METHOD PRIVATE parseFaults : BOOL
VAR
    _q  : UDINT;
    _s  : UDINT;
END_VAR
_q := _device.DCMeter.DCQuesReg;
_s := _swFaultReg;

IF ITECH_Type = 'IT6600C' THEN
    _DeviceFaults.overVoltageProtection  := _q.0;
    _DeviceFaults.overCurrentProtection  := _q.1;
    _DeviceFaults.overPowerProtection    := _q.2;
    _DeviceFaults.underVoltageProtection := _q.3;
    _DeviceFaults.overTempProtection     := _q.4;
    _DeviceFaults.underCurrentProtection := _q.5;
    _DeviceFaults.senseFault             := _q.6;
    _DeviceFaults.currentSharingFault    := _q.7;
    _DeviceFaults.externalInhibit        := _q.9;
    _DeviceFaults.faultProtection        := _q.10;
    _DeviceFaults.loopOscFailure         := _q.11;
    _DeviceFaults.outputNotRegulated     := _q.12;

    _SoftwareFaults.overVoltageProtection         := _s.0;
    _SoftwareFaults.positiveOverCurrentProtection := _s.1;
    _SoftwareFaults.negativeOverCurrentProtection := _s.2;
    _SoftwareFaults.positiveOverPowerProtection   := _s.3;
    _SoftwareFaults.negativeOverPowerProtection   := _s.4;
    _SoftwareFaults.underCurrentProtection        := _s.5;
    _SoftwareFaults.underVoltageProtection        := _s.6;
    _SoftwareFaults.overTemperatureProtection     := _s.7;
END_IF

IF ITECH_Type = 'IT6000' THEN
    _DeviceFaults.overVoltageProtection  := _q.0;
    _DeviceFaults.overCurrentProtection  := _q.1 OR _q.2;
    _DeviceFaults.overPowerProtection    := _q.3 OR _q.4;
    _DeviceFaults.underVoltageProtection := _q.5;
    _DeviceFaults.overTempProtection     := _q.6;
    _DeviceFaults.underCurrentProtection := _q.7;
    _DeviceFaults.senseFault             := _q.8;
    _DeviceFaults.currentSharingFault    := _q.9;
    // bit 10: output reversed (reported through the software-fault register instead)
    _DeviceFaults.externalInhibit        := _q.11;
    _DeviceFaults.faultProtection        := _q.12;
    _DeviceFaults.loopOscFailure         := _q.13;
END_IF

_SoftwareFaults.senseAbnormal                     := _s.8;
_SoftwareFaults.senseReverseProtection            := _s.9;
_SoftwareFaults.outputReverseProtection           := _s.10;
_SoftwareFaults.multiMasterUnitsAbnormal          := _s.11;
_SoftwareFaults.opticalFiberUnlocked_multiMaster  := _s.12;
_SoftwareFaults.opticalFiberUnlocked_singleMaster := _s.13;
_SoftwareFaults.moduleCheckingFailure             := _s.14;
_SoftwareFaults.unevenCurrentProtection           := _s.15;
_SoftwareFaults.hardwareProtection                := _s.16;
_SoftwareFaults.masterUnitPowerFailureProtection  := _s.17;
_SoftwareFaults.inhibit_latchmode                 := _s.18;
_SoftwareFaults.inhibit_livingMode                := _s.19;
_SoftwareFaults.capacitorOverCurrentprotection    := _s.20;
_SoftwareFaults.slaveUnitPowerFailureProtection   := _s.21;
END_METHOD

METHOD PRIVATE rdReal : REAL
VAR_INPUT
    inpIdx      : UINT;
    inpKeep     : REAL;     // returned unchanged unless this signal's last read was good
END_VAR
IF inpIdx <= _readCount AND _arrReadResults[inpIdx].quality = E_SignalQuality.Good THEN
    rdReal := _arrReadResults[inpIdx].valueReal;
ELSE
    rdReal := inpKeep;
END_IF
END_METHOD

METHOD PRIVATE rdUdint : UDINT
VAR_INPUT
    inpIdx      : UINT;
    inpKeep     : UDINT;
END_VAR
IF inpIdx <= _readCount AND _arrReadResults[inpIdx].quality = E_SignalQuality.Good THEN
    rdUdint := _arrReadResults[inpIdx].valueUdint;
ELSE
    rdUdint := inpKeep;
END_IF
END_METHOD

METHOD PRIVATE readImage : BOOL
_device.DCMeter.DCVrms     := rdReal(cRD_METER + 1, _device.DCMeter.DCVrms);
_device.DCMeter.DCIrms     := rdReal(cRD_METER + 2, _device.DCMeter.DCIrms);
_device.DCMeter.DCPrms     := rdReal(cRD_METER + 3, _device.DCMeter.DCPrms);
_device.DCMeter.DCOperReg  := rdUdint(cRD_METER + 4, _device.DCMeter.DCOperReg);
_device.DCMeter.DCStateReg := rdUdint(cRD_METER + 5, _device.DCMeter.DCStateReg);
_device.DCMeter.DCQuesReg  := rdUdint(cRD_METER + 6, _device.DCMeter.DCQuesReg);

_device.DCSource.DCMode          := rdUdint(cRD_SOURCE + 1,  _device.DCSource.DCMode);
_device.DCSource.DCVoltSP        := rdReal(cRD_SOURCE + 2,   _device.DCSource.DCVoltSP);
_device.DCSource.DCVoltRise      := rdReal(cRD_SOURCE + 3,   _device.DCSource.DCVoltRise);
_device.DCSource.DCVoltFall      := rdReal(cRD_SOURCE + 4,   _device.DCSource.DCVoltFall);
_device.DCSource.DCCurrentSP     := rdReal(cRD_SOURCE + 5,   _device.DCSource.DCCurrentSP);
_device.DCSource.DCCurrentRise   := rdReal(cRD_SOURCE + 6,   _device.DCSource.DCCurrentRise);
_device.DCSource.DCCurrentFall   := rdReal(cRD_SOURCE + 7,   _device.DCSource.DCCurrentFall);
_device.DCSource.DCVoltHigh      := rdReal(cRD_SOURCE + 8,   _device.DCSource.DCVoltHigh);
_device.DCSource.DCVoltLow       := rdReal(cRD_SOURCE + 9,   _device.DCSource.DCVoltLow);
_device.DCSource.DCCurrentHigh   := rdReal(cRD_SOURCE + 10,  _device.DCSource.DCCurrentHigh);
_device.DCSource.DCCurrentLow    := rdReal(cRD_SOURCE + 11,  _device.DCSource.DCCurrentLow);
_device.DCSource.DCCC_SpeedState := rdUdint(cRD_SOURCE + 12, _device.DCSource.DCCC_SpeedState);
_device.DCSource.DCCV_SpeedState := rdUdint(cRD_SOURCE + 13, _device.DCSource.DCCV_SpeedState);
_device.DCSource.DCPowerHigh     := rdReal(cRD_SOURCE + 14,  _device.DCSource.DCPowerHigh);
_device.DCSource.DCPowerLow      := rdReal(cRD_SOURCE + 15,  _device.DCSource.DCPowerLow);

_device.Protection.OVPState  := rdUdint(cRD_PROT + 1,  _device.Protection.OVPState);
_device.Protection.OVPLevel  := rdReal(cRD_PROT + 2,   _device.Protection.OVPLevel);
_device.Protection.OVPDelay  := rdReal(cRD_PROT + 3,   _device.Protection.OVPDelay);
_device.Protection.OCPState  := rdUdint(cRD_PROT + 4,  _device.Protection.OCPState);
_device.Protection.OCPLevel  := rdReal(cRD_PROT + 5,   _device.Protection.OCPLevel);
_device.Protection.OCPDelay  := rdReal(cRD_PROT + 6,   _device.Protection.OCPDelay);
_device.Protection.OPPState  := rdUdint(cRD_PROT + 7,  _device.Protection.OPPState);
_device.Protection.OPPLevel  := rdReal(cRD_PROT + 8,   _device.Protection.OPPLevel);
_device.Protection.OPPDelay  := rdReal(cRD_PROT + 9,   _device.Protection.OPPDelay);
_device.Protection.UCPState  := rdUdint(cRD_PROT + 10, _device.Protection.UCPState);
_device.Protection.UCPLevel  := rdReal(cRD_PROT + 11,  _device.Protection.UCPLevel);
_device.Protection.UCPDelay  := rdReal(cRD_PROT + 12,  _device.Protection.UCPDelay);
_device.Protection.UCPWarmup := rdReal(cRD_PROT + 13,  _device.Protection.UCPWarmup);
_device.Protection.UVPState  := rdUdint(cRD_PROT + 14, _device.Protection.UVPState);
_device.Protection.UVPLevel  := rdReal(cRD_PROT + 15,  _device.Protection.UVPLevel);
_device.Protection.UVPDelay  := rdReal(cRD_PROT + 16,  _device.Protection.UVPDelay);
_device.Protection.UVPWarmup := rdReal(cRD_PROT + 17,  _device.Protection.UVPWarmup);

_swFaultReg := rdUdint(cRD_SWF, _swFaultReg);

_device.System.ON_OFF            := rdUdint(cRD_SYS + 1, _device.System.ON_OFF);
_device.System.SenseVolt         := rdReal(cRD_SYS + 2,  _device.System.SenseVolt);
_device.System.Heartbeat         := rdUdint(cRD_SYS + 3, _device.System.Heartbeat);
_device.System.Timer_ON_OFF      := rdUdint(cRD_SYS + 4, _device.System.Timer_ON_OFF);
_device.System.RemoteSenseStatus := rdUdint(cRD_SYS + 5, _device.System.RemoteSenseStatus);
_device.System.RemoteSenseLevel  := rdReal(cRD_SYS + 6,  _device.System.RemoteSenseLevel);
_device.System.OutputRZero       := rdUdint(cRD_SYS + 7, _device.System.OutputRZero);
_device.System.MeasureCycle      := rdUdint(cRD_SYS + 8, _device.System.MeasureCycle);
END_METHOD

METHOD PRIVATE runComms : BOOL
VAR
    _i      : UINT;
END_VAR
// A reset (rising edge) re-arms comms and queues the supply's own protection reset.
_resetTrig(CLK := _resetCalled);
_resetCalled := FALSE;
IF _resetTrig.Q THEN
    _commFaulted := FALSE;
    _deviceResetPending := TRUE;
END_IF

// A type change while running takes comms down for one scan so the driver re-reads its tables.
_mapChanged := _commRunPrev AND (ITECH_Type <> _activeType);
_commRun := _enabled AND _mapValid AND NOT _commFaulted AND NOT _mapChanged;

IF _commRun AND NOT _commRunPrev THEN
    configureDriver();
    _baselineTaken  := FALSE;
    _lastReadCycles := 0;
    _tonReadWatchdog(IN := FALSE);
END_IF
_commRunPrev := _commRun;

IF _baselineTaken THEN
    writeImage();
END_IF

_mb(
    inpEnable           := _commRun,
    inpHoldWrites       := NOT _baselineTaken,
    inpPtrReadConfig    := ADR(_arrReadConfig),
    inpPtrWriteConfig   := ADR(_arrWriteConfig),
    inpPtrReadResults   := ADR(_arrReadResults),
    inpPtrWriteData     := ADR(_arrWriteData));
_mb.cycle();

IF NOT _commRun THEN
    _tonReadWatchdog(IN := FALSE);
    deviceResetWrite();         // keeps the one-shot driver disabled
    RETURN;
END_IF

// ── the latch: the FIRST failed transaction stops everything ────────────────────────────────
IF _mb.stsError THEN
    latchCommFault('Modbus driver configuration error - comms stopped until reset');
    RETURN;
END_IF
FOR _i := 1 TO _readCount DO
    IF _arrReadResults[_i].quality = E_SignalQuality.BadComm THEN
        latchCommFault('Modbus read failed - comms stopped until reset');
        RETURN;
    END_IF
END_FOR
FOR _i := 1 TO cWR_PROT + 17 DO
    IF _arrWriteData[_i].writeError THEN
        latchCommFault('Modbus write failed - comms stopped until reset');
        RETURN;
    END_IF
END_FOR

// A driver that stops completing read cycles without reporting an error is a fault too.
IF _mb.stsStatus.totalReadCycles <> _lastReadCycles THEN
    _lastReadCycles := _mb.stsStatus.totalReadCycles;
    _tonReadWatchdog(IN := FALSE);
END_IF
_tonReadWatchdog(IN := TRUE, PT := _wdTime);
IF _tonReadWatchdog.Q THEN
    latchCommFault('Modbus read watchdog: no read cycle completed - comms stopped until reset');
    RETURN;
END_IF

readImage();

// First complete, clean read cycle since (re)start: seed the command image from the supply,
// then release writes.
IF NOT _baselineTaken AND _mb.stsStatus.totalReadCycles > 0 THEN
    _command := _device;
    IF _baselineCurrentLimit > 0 THEN
        cmdSetCurrentLimits(currentLimitHigh := _baselineCurrentLimit,
                            currentLimitLow  := -_baselineCurrentLimit);
    END_IF
    initParameters();
    IF _commFaultSeen THEN
        cmdDCSourceEnable(FALSE);       // also zeroes the operator's ON/OFF request
        _commFaultSeen := FALSE;
    END_IF
    _baselineTaken := TRUE;
END_IF

deviceResetWrite();
END_METHOD

METHOD PRIVATE selectRegisterMap : BOOL
_mapValid := TRUE;

IF ITECH_Type = 'IT6600C' THEN
    _regDCMeter         := 1401;
    _regDCSource        := 1201;
    _regSystemStatus    := 1001;
    _regProtection      := 1701;
    _regSoftwareFaults  := 1803;
    _regOnOff           := 1001;
    _regResetFault      := 1801;
    _scanTime           := T#100MS;
    _hasExtStatus       := TRUE;
ELSIF ITECH_Type = 'IT6000' THEN
    _regDCMeter         := 1107;
    _regDCSource        := 1019;
    _regSystemStatus    := 1001;
    _regProtection      := 1169;
    _regSoftwareFaults  := 1225;
    _regOnOff           := 1001;
    _regResetFault      := 1223;
    _scanTime           := T#250MS;
    _hasExtStatus       := FALSE;
ELSE
    _mapValid := FALSE;
END_IF
END_METHOD

METHOD setCommandValues : BOOL
IF NOT inpAuto THEN
    IF NOT stsFaulted THEN
        _command.System.ON_OFF     := HMI_DeviceSignals.deviceSignals_write.System.ON_OFF;
        _command.DCSource.DCMode   := HMI_DeviceSignals.deviceSignals_write.DCSource.DCMode;
    END_IF
    _command.DCSource.DCPowerHigh   := HMI_DeviceSignals.deviceSignals_write.DCSource.DCPowerHigh;
    _command.DCSource.DCPowerLow    := HMI_DeviceSignals.deviceSignals_write.DCSource.DCPowerLow;
    _command.DCSource.DCCurrentSP   := HMI_DeviceSignals.deviceSignals_write.DCSource.DCCurrentSP;
    _command.DCSource.DCCurrentRise := HMI_DeviceSignals.deviceSignals_write.DCSource.DCCurrentRise;
    _command.DCSource.DCCurrentFall := HMI_DeviceSignals.deviceSignals_write.DCSource.DCCurrentFall;
    _command.DCSource.DCCurrentHigh := HMI_DeviceSignals.deviceSignals_write.DCSource.DCCurrentHigh;
    _command.DCSource.DCCurrentLow  := HMI_DeviceSignals.deviceSignals_write.DCSource.DCCurrentLow;
    _command.DCSource.DCVoltSP      := HMI_DeviceSignals.deviceSignals_write.DCSource.DCVoltSP;
    _command.DCSource.DCVoltRise    := HMI_DeviceSignals.deviceSignals_write.DCSource.DCVoltRise;
    _command.DCSource.DCVoltFall    := HMI_DeviceSignals.deviceSignals_write.DCSource.DCVoltFall;
    _command.DCSource.DCVoltHigh    := HMI_DeviceSignals.deviceSignals_write.DCSource.DCVoltHigh;
    _command.DCSource.DCVoltLow     := HMI_DeviceSignals.deviceSignals_write.DCSource.DCVoltLow;

    _command.Protection.OCPState    := HMI_DeviceSignals.deviceSignals_write.Protection.OCPState;
    _command.Protection.OCPLevel    := HMI_DeviceSignals.deviceSignals_write.Protection.OCPLevel;
    _command.Protection.OCPDelay    := HMI_DeviceSignals.deviceSignals_write.Protection.OCPDelay;
    _command.Protection.OVPState    := HMI_DeviceSignals.deviceSignals_write.Protection.OVPState;
    _command.Protection.OVPLevel    := HMI_DeviceSignals.deviceSignals_write.Protection.OVPLevel;
    _command.Protection.OVPDelay    := HMI_DeviceSignals.deviceSignals_write.Protection.OVPDelay;
    _command.Protection.UCPState    := HMI_DeviceSignals.deviceSignals_write.Protection.UCPState;
    _command.Protection.UCPLevel    := HMI_DeviceSignals.deviceSignals_write.Protection.UCPLevel;
    _command.Protection.UCPDelay    := HMI_DeviceSignals.deviceSignals_write.Protection.UCPDelay;
    _command.Protection.UVPState    := HMI_DeviceSignals.deviceSignals_write.Protection.UVPState;
    _command.Protection.UVPLevel    := HMI_DeviceSignals.deviceSignals_write.Protection.UVPLevel;
    _command.Protection.UVPDelay    := HMI_DeviceSignals.deviceSignals_write.Protection.UVPDelay;
    _command.Protection.OPPState    := HMI_DeviceSignals.deviceSignals_write.Protection.OPPState;
    _command.Protection.OPPLevel    := HMI_DeviceSignals.deviceSignals_write.Protection.OPPLevel;
    _command.Protection.OPPDelay    := HMI_DeviceSignals.deviceSignals_write.Protection.OPPDelay;
END_IF
END_METHOD

METHOD setConfigs : BOOL
VAR_INPUT
    configs : ST_ITECH_SetConfigs;
END_VAR
_command.DCSource.DCMode         := configs.dcSource.DCMode;
_command.DCSource.DCPowerHigh    := configs.dcSource.DCPowerHigh;
_command.DCSource.DCPowerLow     := configs.dcSource.DCPowerLow;
_command.DCSource.DCCurrentSP    := configs.dcSource.DCCurrentSP;
_command.DCSource.DCCurrentRise  := configs.dcSource.DCCurrentRise;
_command.DCSource.DCCurrentFall  := configs.dcSource.DCCurrentFall;
_command.DCSource.DCCurrentHigh  := configs.dcSource.DCCurrentHigh;
_command.DCSource.DCCurrentLow   := configs.dcSource.DCCurrentLow;
_command.DCSource.DCVoltSP       := configs.dcSource.DCVoltSP;
_command.DCSource.DCVoltRise     := configs.dcSource.DCVoltRise;
_command.DCSource.DCVoltFall     := configs.dcSource.DCVoltFall;
_command.DCSource.DCVoltHigh     := configs.dcSource.DCVoltHigh;
_command.DCSource.DCVoltLow      := configs.dcSource.DCVoltLow;

_command.Protection.OCPLevel     := configs.protection.OCPLevel;
_command.Protection.OCPDelay     := configs.protection.OCPDelay;
_command.Protection.UCPLevel     := configs.protection.UCPLevel;
_command.Protection.UCPDelay     := configs.protection.UCPDelay;
_command.Protection.OVPLevel     := configs.protection.OVPLevel;
_command.Protection.OVPDelay     := configs.protection.OVPDelay;
_command.Protection.UVPLevel     := configs.protection.UVPLevel;
_command.Protection.UVPDelay     := configs.protection.UVPDelay;
_command.Protection.OPPLevel     := configs.protection.OPPLevel;
_command.Protection.OPPDelay     := configs.protection.OPPDelay;

_command.Protection.UCPState     := configs.protection.UCPState;
_command.Protection.UVPState     := configs.protection.UVPState;
_command.Protection.OCPState     := configs.protection.OCPState;
_command.Protection.OVPState     := configs.protection.OVPState;
_command.Protection.OPPState     := configs.protection.OPPState;
END_METHOD

METHOD setInterlock : BOOL
Interlock.name := _DeviceName;
Interlock(inpConfig := _dataInterlock);
END_METHOD

METHOD PRIVATE setRead : BOOL
VAR_INPUT
    inpIdx      : UINT;
    inpReg      : UINT;     // protocol (0-based) holding-register address
    inpIsReal   : BOOL;     // TRUE = 32-bit float, FALSE = 32-bit unsigned
END_VAR
_arrReadConfig[inpIdx].modbusAddr := 400001 + UINT_TO_UDINT(inpReg);
IF inpIsReal THEN
    _arrReadConfig[inpIdx].dataType := E_MBDataType.mbReal32;
ELSE
    _arrReadConfig[inpIdx].dataType := E_MBDataType.mbUInt32;
END_IF
END_METHOD

METHOD setStatusValues : BOOL
stsDCSourceState := _device.System.ON_OFF;
stsDCMode        := _device.DCSource.DCMode;
stsDCSource_V_SP := _device.DCSource.DCVoltSP;
stsDCMeterV      := _device.DCMeter.DCVrms;
stsDCMeterI      := _device.DCMeter.DCIrms;
stsDCMeterP      := _device.DCMeter.DCPrms;
sendLog(CONCAT('DC Source state changed to ', TO_STRING(stsDCSourceState)), 1);
sendLog(CONCAT('DC Source Voltage setpoint set to ', TO_STRING(stsDCSource_V_SP)), 2);
sendLog(CONCAT('DC Source mode set to ', TO_STRING(stsDCMode)), 3);
END_METHOD

METHOD PRIVATE setWrite : BOOL
VAR_INPUT
    inpIdx      : UINT;
    inpReg      : UINT;
    inpIsReal   : BOOL;
END_VAR
_arrWriteConfig[inpIdx].modbusAddr := 400001 + UINT_TO_UDINT(inpReg);
IF inpIsReal THEN
    _arrWriteConfig[inpIdx].dataType := E_MBDataType.mbReal32;
ELSE
    _arrWriteConfig[inpIdx].dataType := E_MBDataType.mbUInt32;
END_IF
END_METHOD

METHOD PRIVATE updateHMI : BOOL
HMI_DeviceSignals.deviceSignals_read := _device;
END_METHOD

METHOD PRIVATE writeImage : BOOL
// ON/OFF goes out as two 16-bit registers, LOW word first — exactly the bytes the previous
// implementation sent (it wrote the raw UDINT, not the word-swapped image every other value
// uses). Kept byte-for-byte because the supplies run on it; it is the one asymmetry with the
// read side (which takes the register pair high word first), so verify against the supply's
// manual before "fixing" it.
_arrWriteData[cWR_ONOFF + 1].valueUint := UDINT_TO_UINT(_command.System.ON_OFF AND 16#FFFF);
_arrWriteData[cWR_ONOFF + 2].valueUint := UDINT_TO_UINT(SHR(_command.System.ON_OFF, 16));

// IT6000 power values are in kW, IT6600C power values in W
_arrWriteData[cWR_SOURCE + 1].valueUdint := _command.DCSource.DCMode;
_arrWriteData[cWR_SOURCE + 2].valueReal  := _command.DCSource.DCVoltSP;
_arrWriteData[cWR_SOURCE + 3].valueReal  := _command.DCSource.DCVoltRise;
_arrWriteData[cWR_SOURCE + 4].valueReal  := _command.DCSource.DCVoltFall;
_arrWriteData[cWR_SOURCE + 5].valueReal  := _command.DCSource.DCCurrentSP;
_arrWriteData[cWR_SOURCE + 6].valueReal  := _command.DCSource.DCCurrentRise;
_arrWriteData[cWR_SOURCE + 7].valueReal  := _command.DCSource.DCCurrentFall;
_arrWriteData[cWR_SOURCE + 8].valueReal  := _command.DCSource.DCVoltHigh;
_arrWriteData[cWR_SOURCE + 9].valueReal  := _command.DCSource.DCVoltLow;
_arrWriteData[cWR_SOURCE + 10].valueReal := _command.DCSource.DCCurrentHigh;
_arrWriteData[cWR_SOURCE + 11].valueReal := _command.DCSource.DCCurrentLow;
_arrWriteData[cWR_SOURCE + 12].valueUdint := _command.DCSource.DCCC_SpeedState;
_arrWriteData[cWR_SOURCE + 13].valueUdint := _command.DCSource.DCCV_SpeedState;
_arrWriteData[cWR_SOURCE + 14].valueReal := _command.DCSource.DCPowerHigh;
_arrWriteData[cWR_SOURCE + 15].valueReal := _command.DCSource.DCPowerLow;

_arrWriteData[cWR_PROT + 1].valueUdint  := _command.Protection.OVPState;
_arrWriteData[cWR_PROT + 2].valueReal   := _command.Protection.OVPLevel;
_arrWriteData[cWR_PROT + 3].valueReal   := _command.Protection.OVPDelay;
_arrWriteData[cWR_PROT + 4].valueUdint  := _command.Protection.OCPState;
_arrWriteData[cWR_PROT + 5].valueReal   := _command.Protection.OCPLevel;
_arrWriteData[cWR_PROT + 6].valueReal   := _command.Protection.OCPDelay;
_arrWriteData[cWR_PROT + 7].valueUdint  := _command.Protection.OPPState;
_arrWriteData[cWR_PROT + 8].valueReal   := _command.Protection.OPPLevel;
_arrWriteData[cWR_PROT + 9].valueReal   := _command.Protection.OPPDelay;
_arrWriteData[cWR_PROT + 10].valueUdint := _command.Protection.UCPState;
_arrWriteData[cWR_PROT + 11].valueReal  := _command.Protection.UCPLevel;
_arrWriteData[cWR_PROT + 12].valueReal  := _command.Protection.UCPDelay;
_arrWriteData[cWR_PROT + 13].valueReal  := _command.Protection.UCPWarmup;
_arrWriteData[cWR_PROT + 14].valueUdint := _command.Protection.UVPState;
_arrWriteData[cWR_PROT + 15].valueReal  := _command.Protection.UVPLevel;
_arrWriteData[cWR_PROT + 16].valueReal  := _command.Protection.UVPDelay;
_arrWriteData[cWR_PROT + 17].valueReal  := _command.Protection.UVPWarmup;
END_METHOD

END_FUNCTION_BLOCK

// ---- POUs/FBs/Devices/fb_Dev_Pump_SPAL.TcPOU
FUNCTION_BLOCK fb_Dev_Pump_SPAL EXTENDS abs_fb_Device
VAR_INPUT
	IO_CANIn		: POINTER TO ST_Pump_SPAL_CAN_Inputs;
	IO_CANOut		: POINTER TO ST_Pump_SPAL_CAN_Outputs;
	IO_CAN_State	: POINTER TO ST_EL6751_Bus_State;
	IO_LV_DO		: POINTER TO BOOL;
	inpESTOPActive	: BOOL;
	inpMachineSTOP	: BOOL;
END_VAR

VAR PERSISTENT
	HMI						: ST_Pump_SPAL_HMI_Interface;
END_VAR
	
VAR
	LVActuator				:fb_Dev_Actuator(cfgDeviceName := CONCAT(_deviceName,' PWR'), cfgHasFeedback:=FALSE,cfgInitEventclass := TRUE,
										  cfgEnable := TRUE,
										  cfgOnDelay :=T#3S,
										  cfgOffDelay:=T#1S,
										  cfgRetractOnFault := TRUE,
										  cfgInvFeedback:=FALSE);
	_LVActuator_interlocks	: ARRAY [1..10] OF BOOL;
	_interlocks				: ARRAY [1..10] of BOOL;
	
	Bus_Status				: fb_IO_EL6751_Bus_Status;
	_pumpState				: STRING;
	_pumpCommandFB			: STRING;
	_pumpMotorFB			: STRING;
	_pumpServiceIndicator	: STRING;
	_pumpError				: STRING;
	_pumpPower				: LREAL;
	_pumpTemperature		: LREAL;
	_pumpSpeed				: LREAL;
	_ctrlRunPump			: USINT;
	_ctrlSetpoint			: LREAL;
END_VAR

VAR_OUTPUT
	stsLVOn		: BOOL;
	stsEnabled	: BOOL;
END_VAR

DeviceLogic();
Bus_Status(IO_Bus_State	:= IO_CAN_State^);
LVActuator(inpAuto:= inpAuto,inpReset:=inpReset,IO_output_Actuate:=IO_LV_DO^);

_LVActuator_interlocks[1] := inpESTOPActive;
LVActuator.cmdSetInterlock(1,'ESTOPs Not Active',_LVActuator_interlocks[1]);

_interlocks[1] := inpESTOPActive;
cmdSetInterlock(1,'ESTOPs Not Active',_LVActuator_interlocks[1]);

_interlocks[2] := LVactuator.stsActuated;
cmdSetInterlock(2, 'LV On', _interlocks[2]);

_interlocks[3] := NOT(inpMachineStop);
cmdSetInterlock(3, 'Machine STOP Not Active', _interlocks[3]);


parsePumpFeedback();
FaultHandler();

IF _Enabled THEN
	IF (NOT _inAuto) THEN
		_ctrlRunPump	:= HMI.ocmdRunPump;
		_ctrlSetpoint	:= HMI.ocmdSetpoint;
	END_IF
END_IF

IF NOT(LVActuator.stsActuated) THEN
	resetControlSignals();
END_IF

// A faulted pump is not commanded to run. Without this, an auto-mode run request survived the
// fault and the pump restarted by itself as soon as its interlock came back.
IF stsFaulted THEN
	_ctrlRunPump    := 0;
	HMI.ocmdRunPump := 0;
END_IF

IF interlock.outInterlockOK THEN
	IO_CANOut^.MotorSetpoint 	:= _ctrlSetpoint;
	IO_CANOut^.MotorStateRequest := _ctrlRunPump;
ELSE
	HMI.ocmdRunPump := 0;
	IO_CANOut^.MotorStateRequest := 0;
END_IF

sendLog(Concat('Run command set to ',TO_STRING(_ctrlRunPump)),1);
sendLog(Concat('Setpoint set to ', TO_STRING(_ctrlSetpoint)),2);

updateHMI();

stsLVOn	:= LVActuator.stsActuated;
stsEnabled := (_ctrlRunPump = 1);

METHOD cmdEnable : BOOL
VAR_INPUT
	command	: USINT; //1= Enable, 0= Disable
END_VAR
_ctrlRunPump := command;
END_METHOD

METHOD PUBLIC cmdLV : BOOL
VAR_INPUT
	command	: BOOL; //1=ON, 0=OFF
END_VAR
IF command THEN
	LVActuator.cmdActuate();
ELSE
	LVActuator.cmdRetract();
END_IF
END_METHOD

METHOD cmdReset : BOOL
setFault(0,'');
END_METHOD

METHOD cmdSetpoint : BOOL
VAR_INPUT
	setpoint	: LREAL; //0-100%
END_VAR
_ctrlSetpoint	:= setpoint;
END_METHOD

METHOD PRIVATE FaultHandler : BOOL
VAR_INPUT
END_VAR


IF LVActuator.stsFaulted AND _ctrlRunPump = 1 THEN
	setFault(1,LVActuator.stsFaultDescription);
END_IF

IF LVactuator.stsActuated AND _ctrlRunPump = 1 AND IO_CANIn^.PumpOperatorStatus = EN_Pump_SPAL_Operating_status.Not_Operable THEN 
	setFault(1,_pumpError);
END_IF

// Faults LATCH until cmdReset / inpReset. (A 'Normal' operating status used to clear every fault
// here on the next scan, interlock-loss and LV faults included, so nothing stayed faulted.)

IF IO_CANIn^.PumpOperatorStatus = EN_Pump_SPAL_Operating_status.Derated THEN
	sendWarning('Derated',10);
END_IF

IF IO_CANIn^.PumpServiceIndicator = EN_Pump_SPAL_ServiceIndicator.Service_required THEN
	sendWarning('Service required',11);
END_IF

//If enabled and  then fault
IF NOT stsFaulted AND _ctrlRunPump = 1 THEN
	IF NOT interlock.outInterlockOK THEN
		setFault(1,CONCAT('I_NOK - ',Interlock.stsFirstOut));
	END_IF
END_IF
END_METHOD

//FB_Init is always available implicitly and it is used primarily for initialization.
//The return value is not evaluated. For a specific influence, you can also declare the
//methods explicitly and provide additional code there with the standard initialization
//code. You can evaluate the return value.
METHOD FB_Init: BOOL
VAR_INPUT
    bInitRetains: BOOL; // TRUE: the retain variables are initialized (reset warm / reset cold)
    bInCopyCode: BOOL;  // TRUE: the instance will be copied to the copy code afterward (online change) 
	cfgDeviceName 	: STRING;
	cfgEnable		: BOOL;
	cfgInitEventClass	: BOOL;
END_VAR
THIS^.cfgDeviceName 	:= cfgDeviceName;
THIS^.cfgEnable 		:= cfgEnable;
THIS^.cfgInitEventClass	:= cfgInitEventClass;
END_METHOD

METHOD PRIVATE parsePumpFeedback : BOOL
VAR_INPUT
END_VAR
CASE TO_INT(IO_CANIn^.PumpError) OF
	EN_Pump_SPAL_PumpError.Dry_Run:
		_pumpError :=   'Dry Run';
	EN_Pump_SPAL_PumpError.Normal_Operation:
		_pumpError := 'N/A';
	EN_Pump_SPAL_PumpError.OverT_Protection_Shutdown:
		_pumpError := 'Over Temperature Protection';
	EN_Pump_SPAL_PumpError.OverV_Protection_Shutdown:
		_pumpError := 'Over Voltage Protection';
	EN_Pump_SPAL_PumpError.Speed_Limited_Due_To_Capability:
		_pumpError := 'Speed limited due to capability';
	EN_Pump_SPAL_PumpError.Speed_Limited_Due_To_Current:
		_pumpError := 'Speed limited due to current';
	EN_Pump_SPAL_PumpError.Speed_Limited_Due_To_OverT:
		_pumpError := 'Speed limited due to overtemperature';
	EN_Pump_SPAL_PumpError.Speed_Limited_Due_To_Torque:
		_pumpError := 'Speed limited due to torque';
	EN_Pump_SPAL_PumpError.Unable_to_start:
		_pumpError := 'Unable to start';
	EN_Pump_SPAL_PumpError.UnderV_Protection_Shutdown:
		_pumpError := 'Undervoltage protection';
	ELSE
		_pumpError := 'Undefined error';
		
END_CASE

CASE TO_INT(IO_CANIn^.PumpOperatorStatus) OF
	EN_Pump_SPAL_Operating_status.Derated:
		_pumpState := 'Derated';
	EN_Pump_SPAL_Operating_status.Normal:
		_pumpState := 'Normal';
	EN_Pump_SPAL_Operating_status.Not_Available:
		_pumpState := 'Not Available';
	EN_Pump_SPAL_Operating_status.Not_Operable:
		_pumpState:= 'Not Operable';	
END_CASE

CASE TO_INT(IO_CANIn^.PumpServiceIndicator) OF
	EN_Pump_SPAL_ServiceIndicator.Not_Available:
		_pumpServiceIndicator := 'N/A';
	EN_Pump_SPAL_ServiceIndicator.Reserved:
		_pumpServiceIndicator:= 'Reserved';
	EN_Pump_SPAL_ServiceIndicator.Service_not_required:
		_pumpServiceIndicator := 'OK';
	EN_Pump_SPAL_ServiceIndicator.Service_required:
		_pumpServiceIndicator := 'Service Required';	
END_CASE

CASE TO_INT(IO_CANIn^.PumpCMDStatus) OF
	0:
		_pumpCommandFB := 'Internal';
	1:
		_pumpCommandFB := 'External';
	2:
		_pumpCommandFB := 'Default';
	3:
		_pumpCommandFB := 'N/A';
END_CASE

CASE TO_INT(IO_CANIn^.PumpMotor) OF
	0:
		_pumpMotorFB := 'OFF';
	1:
		_pumpMotorFB := 'ON';
	2:
		_pumpMotorFB := 'Reverse';
	3:
		_pumpMotorFB := 'N/A';
END_CASE

_pumpTemperature := IO_CANIn^.PumpTemperature;
_pumpSpeed		 := IO_CANIn^.PumpSpeed;
_pumpPower		 := IO_CANIn^.PumpPower;
END_METHOD

METHOD PRIVATE resetControlSignals : BOOL
VAR_INPUT
END_VAR
_ctrlRunPump	:= 0;
_ctrlSetpoint	:= 0.0;
END_METHOD

METHOD PRIVATE updateHMI : BOOL
VAR

END_VAR
HMI.HMIbaseDevice := HMIbaseDevice;
HMI.stsBusStatus  := Bus_Status.getHMIData();

HMI.stsRunPump	  := _ctrlRunPump;
HMI.stsSetpoint	  := _ctrlSetpoint;

HMI.stsCommandFB 		:= _pumpCommandFB;
HMI.stsError	 		:= _pumpError;
HMI.stsMotorFB			:= _pumpMotorFB;
HMI.stsPower     		:= _pumpPower;
HMI.stsServiceIndicator := _pumpServiceIndicator;
HMI.stsSpeed			:= _pumpSpeed;
HMI.stsState			:= _pumpState;
HMI.stsTemperature		:= _pumpTemperature;

IF bus_status.stsBusFaulted THEN
	HMI.stsBusOK := FALSE;
ELSE
	HMI.stsBusOK := TRUE;
END_IF
END_METHOD

END_FUNCTION_BLOCK

// ---- POUs/FBs/fb_IO_EL6751_Bus_Status.TcPOU
FUNCTION_BLOCK fb_IO_EL6751_Bus_Status
VAR_INPUT
	IO_Bus_State	:	ST_EL6751_Bus_State;
END_VAR
VAR_OUTPUT
	stsBusFaulted	: BOOL;
END_VAR
VAR
	HMI			:ST_EL6751_Bus_State_Parsed;
	_busState	:ST_EL6751_Bus_State_Parsed;	
END_VAR

_busState.stsBusLoad 					:= IO_Bus_State.GlobalState3;


_busState.stsCANControllerBusOff		:= IO_Bus_State.GlobalState2.Bits[1].Bit1;
_busState.stsCANControllerWarningLimit	:= IO_bus_State.GlobalState2.Bits[1].Bit2;
_busState.stsRxQueueOverrun				:= IO_bus_State.GlobalState2.Bits[1].Bit3;
_busState.stsCANSendError				:= IO_bus_State.GlobalState2.Bits[1].Bit6;
_busState.stsCANQueueIntRxOverflow		:= IO_bus_State.GlobalState2.Bits[1].Bit8;
_busState.stsCANQueueIntTxOverflow		:= IO_bus_State.GlobalState2.Bits[1].Bit9;
_busState.stsSyncToggle					:= IO_bus_State.GlobalState2.Bits[1].Bit16;

CASE IO_Bus_State.GlobalState0 OF
	0:
		_busState.stsCANDeviceState	:= 'RUN';
	1:
		_busState.stsCANDeviceState	:= 'RESET';
	2:
		_busState.stsCANDeviceState	:= 'OFFLINE';
	3:
		_busState.stsCANDeviceState	:= 'STOP';
	ELSE
		_busState.stsCANDeviceState	:= 'ERR';
END_CASE

IF (IO_Bus_State.GlobalState0 <> 0) OR (IO_Bus_State.GlobalState2.Num <> 0) THEN
	stsBusFaulted := TRUE;
ELSE
	stsBusFaulted := FALSE;
END_IF

HMI := _busState;

METHOD PUBLIC getHMIData : ST_EL6751_Bus_State_Parsed
VAR_INPUT
END_VAR
getHMIData := HMI;
END_METHOD

END_FUNCTION_BLOCK

// ---- POUs/FBs/Devices/fb_Dev_StackLight3SegHV_BannerTL50Pro.TcPOU
FUNCTION_BLOCK fb_Dev_StackLight3SegHV_BannerTL50Pro
VAR_INPUT
	IOOut_BannerTL503Pro: POINTER TO ST_Banner_TL503Pro_Raw;
	inpFaulted			: BOOL;
	inpSafetyFaultActive: BOOL;
	inpHVOn				: BOOL;
	inpMotionPresent	: BOOL;
	inpAuto				: BOOL;
	inpRunningInAuto	: BOOL;
	inpDoneInAuto		: BOOL;
	
END_VAR

VAR
	_stackLightState	: INT;
	_stackLight			: ST_Banner_TL503Pro;
	
END_VAR

//Constant values
_stackLight.Segment1Color1.Num := TO_USINT(EN_Banner_TL503Pro_Colors.Orange);
_stackLight.Segment2Color2.Num := TO_USINT(EN_Banner_TL503Pro_Colors.Orange);
_stackLight.Segment3Color1.Num := TO_USINT(EN_Banner_TL503Pro_Colors.Red);

//Temp logic for segment2 until state machine exists
IF NOT(inpAuto) THEN
	IF inpMotionPresent  THEN
		_stackLightState := 1;
	ELSE
		_stackLightState := 0;
	END_IF
ELSE
	IF inpRunningInAuto THEN
		IF inpMotionPresent THEN
			_stackLightState := 12;
		ELSE
			_stackLightState := 11;
		END_IF
	ELSE
		IF inpDoneInAuto THEN
			_stackLightState := 20;
		ELSE
			_stackLightState := 10;
		END_IF
	END_IF
END_IF

IF inpHVOn THEN
	_stackLight.Segment1AnimationType.Num 		:= TO_USINT(EN_Banner_TL503Pro_Animation.Steady);
ELSE
	_stackLight.Segment1AnimationType.Num 		:= TO_USINT(EN_Banner_TL503Pro_Animation.Off);
END_IF

IF inpFaulted THEN
	_stackLight.Segment3AnimationType.Num 		:= TO_USINT(EN_Banner_TL503Pro_Animation.Steady);
END_IF

IF inpSafetyFaultActive THEN
	_stackLight.Segment3AnimationType.Num 		:= TO_USINT(EN_Banner_TL503Pro_Animation.IntensitySweep);
END_IF

IF (NOT inpFaulted) AND (NOT inpSafetyFaultActive) THEN
	_stackLight.Segment3AnimationType.Num 		:= TO_USINT(EN_Banner_TL503Pro_Animation.off);
END_IF

CASE _stackLightState OF
    0:
    // Manual, Not running    
        _stackLight.Segment2Color1.Num 			:= TO_USINT(EN_Banner_TL503Pro_Colors.White);
        _stackLight.Segment2AnimationType.Num 	:= TO_USINT(EN_Banner_TL503Pro_Animation.Steady);
    1:
    // Manual, Motion
        _stackLight.Segment2Color1.Num 			:= TO_USINT(EN_Banner_TL503Pro_Colors.White);
        _stackLight.Segment2AnimationType.Num 	:= TO_USINT(EN_Banner_TL503Pro_Animation.FiftyFiftyRotate);
	2:
	//Manual, coolant but no motion
		_stackLight.Segment2Color1.Num 			:= TO_USINT(EN_Banner_TL503Pro_Colors.White);
		_stackLight.Segment2Color2.Num 			:= TO_USINT(EN_Banner_TL503Pro_Colors.Blue);
		_stackLight.Segment2AnimationType.Num 	:= TO_USINT(EN_Banner_TL503Pro_Animation.Chase);
    10:
    // Auto, Not Running, No Motion
        _stackLight.Segment2Color1.Num 			:= TO_USINT(EN_Banner_TL503Pro_Colors.Green);
        _stackLight.Segment2AnimationType.Num 	:= TO_USINT(EN_Banner_TL503Pro_Animation.IntensitySweep);
    11:
	// Auto, Running, No Motion
        _stackLight.Segment2Color1.Num 			:= TO_USINT(EN_Banner_TL503Pro_Colors.Green);
        _stackLight.Segment2AnimationType.Num 	:= TO_USINT(EN_Banner_TL503Pro_Animation.Steady);

    12:
    // Auto, Running, Motion
        // (Segment 1 is the HV indicator and is driven ONLY by inpHVOn above. This state used to
        // force it on, so the light showed HV ON with HV off whenever the machine ran in auto.)
        _stackLight.Segment2Color1.Num 			:= TO_USINT(EN_Banner_TL503Pro_Colors.Green);
        _stackLight.Segment2AnimationType.Num 	:= TO_USINT(EN_Banner_TL503Pro_Animation.FiftyFiftyRotate);
		
	20:
	//Auto, Done
		_stackLight.Segment2Color1.Num 			:= TO_USINT(EN_Banner_TL503Pro_Colors.Blue);
        _stackLight.Segment2AnimationType.Num 	:= TO_USINT(EN_Banner_TL503Pro_Animation.IntensitySweep);

	ELSE
	// Unknown state: flash segment 2 blue. Segment 1 (HV) is never repurposed.
		_stackLight.Segment2Color1.Num 			:= TO_USINT(EN_Banner_TL503Pro_Colors.Blue);
		_stackLight.Segment2AnimationType.Num 	:= TO_USINT(EN_Banner_TL503Pro_Animation.Flash);

END_CASE

writeToPDO(_stackLight,IOOut_BannerTL503Pro);

METHOD PRIVATE writeToPDO : BOOL
VAR_INPUT
	SignalArray : ST_Banner_TL503Pro;
	OutputArray : POINTER TO ST_Banner_TL503Pro_Raw;
END_VAR
//Segment1 Color1
OutputArray^.PDOs[30].0 := SignalArray.Segment1Color1.Bits[1].Bit1;
OutputArray^.PDOs[30].1 := SignalArray.Segment1Color1.Bits[1].Bit2;
OutputArray^.PDOs[30].2 := SignalArray.Segment1Color1.Bits[1].Bit3;
OutputArray^.PDOs[30].3 := SignalArray.Segment1Color1.Bits[1].Bit4;

//Segment1 Color Intensity
OutputArray^.PDOs[30].4 := SignalArray.Segment1Color1Intensity.Bits[1].Bit1;
OutputArray^.PDOs[30].5 := SignalArray.Segment1Color1Intensity.Bits[1].Bit2;
OutputArray^.PDOs[30].6 := SignalArray.Segment1Color1Intensity.Bits[1].Bit3;
OutputArray^.PDOs[30].7 := SignalArray.Segment1Color1Intensity.Bits[1].Bit4;

//Segment1 Animation Type
OutputArray^.PDOs[29].0 := SignalArray.Segment1AnimationType.Bits[1].Bit1;
OutputArray^.PDOs[29].1 := SignalArray.Segment1AnimationType.Bits[1].Bit2;
OutputArray^.PDOs[29].2 := SignalArray.Segment1AnimationType.Bits[1].Bit3;

//Segment1 Speed
OutputArray^.PDOs[29].3 := SignalArray.Segment1Speed.Bits[1].Bit1;
OutputArray^.PDOs[29].4 := SignalArray.Segment1Speed.Bits[1].Bit2;

//Segment1 Pulse Pattern
OutputArray^.PDOs[29].5 := SignalArray.Segment1PulsePattern.Bits[1].Bit1;
OutputArray^.PDOs[29].6 := SignalArray.Segment1PulsePattern.Bits[1].Bit2;

//Segment1 Color2
OutputArray^.PDOs[28].0 := SignalArray.Segment1Color2.Bits[1].Bit1;
OutputArray^.PDOs[28].1 := SignalArray.Segment1Color2.Bits[1].Bit2;
OutputArray^.PDOs[28].2 := SignalArray.Segment1Color2.Bits[1].Bit3;
OutputArray^.PDOs[28].3 := SignalArray.Segment1Color2.Bits[1].Bit4;

//Segment1 Color2 Intensity
OutputArray^.PDOs[28].4 := SignalArray.Segment1Color2Intensity.Bits[1].Bit1;
OutputArray^.PDOs[28].5 := SignalArray.Segment1Color2Intensity.Bits[1].Bit2;
OutputArray^.PDOs[28].6 := SignalArray.Segment1Color2Intensity.Bits[1].Bit3;

//Segment1 Rotate
OutputArray^.PDOs[28].7 := SignalArray.Segment1RotationDir;

//Segment2 Color1
OutputArray^.PDOs[27].0 := SignalArray.Segment2Color1.Bits[1].Bit1;
OutputArray^.PDOs[27].1 := SignalArray.Segment2Color1.Bits[1].Bit2;
OutputArray^.PDOs[27].2 := SignalArray.Segment2Color1.Bits[1].Bit3;
OutputArray^.PDOs[27].3 := SignalArray.Segment2Color1.Bits[1].Bit4;

//Segment2 Color1 Intensity
OutputArray^.PDOs[27].4 := SignalArray.Segment2Color1Intensity.Bits[1].Bit1;
OutputArray^.PDOs[27].5 := SignalArray.Segment2Color1Intensity.Bits[1].Bit2;
OutputArray^.PDOs[27].6 := SignalArray.Segment2Color1Intensity.Bits[1].Bit3;

//Segment2 Animation Type
OutputArray^.PDOs[26].0 := SignalArray.Segment2AnimationType.Bits[1].Bit1;
OutputArray^.PDOs[26].1 := SignalArray.Segment2AnimationType.Bits[1].Bit2;
OutputArray^.PDOs[26].2 := SignalArray.Segment2AnimationType.Bits[1].Bit3;

//Segment2 Speed
OutputArray^.PDOs[26].3 := SignalArray.Segment2Speed.Bits[1].Bit1;
OutputArray^.PDOs[26].4 := SignalArray.Segment2Speed.Bits[1].Bit2;

//Segment2 Pulse Pattern
OutputArray^.PDOs[26].5 := SignalArray.Segment2PulsePattern.Bits[1].Bit1;
OutputArray^.PDOs[26].6 := SignalArray.Segment2PulsePattern.Bits[1].Bit2;

//Segment 2 Color 2
OutputArray^.PDOs[25].0 := SignalArray.Segment2Color2.Bits[1].Bit1;
OutputArray^.PDOs[25].1 := SignalArray.Segment2Color2.Bits[1].Bit2;
OutputArray^.PDOs[25].2 := SignalArray.Segment2Color2.Bits[1].Bit3;
OutputArray^.PDOs[25].3 := SignalArray.Segment2Color2.Bits[1].Bit4;

//Segment 2 Color 2 Intensity
OutputArray^.PDOs[25].4 := SignalArray.Segment2Color2Intensity.Bits[1].Bit1;
OutputArray^.PDOs[25].5 := SignalArray.Segment2Color2Intensity.Bits[1].Bit2;
OutputArray^.PDOs[25].6 := SignalArray.Segment2Color2Intensity.Bits[1].Bit3;

//Segment 2 Rotate
OutputArray^.PDOs[25].7 := SignalArray.Segment2RotationDir;

//Segment 3 Color 1
OutputArray^.PDOs[24].0 := SignalArray.Segment3Color1.Bits[1].Bit1;
OutputArray^.PDOs[24].1 := SignalArray.Segment3Color1.Bits[1].Bit2;
OutputArray^.PDOs[24].2 := SignalArray.Segment3Color1.Bits[1].Bit3;
OutputArray^.PDOs[24].3 := SignalArray.Segment3Color1.Bits[1].Bit4;

//Segment 3 Color1 Intensity
OutputArray^.PDOs[24].4 := SignalArray.Segment3Color1Intensity.Bits[1].Bit1;
OutputArray^.PDOs[24].5 := SignalArray.Segment3Color1Intensity.Bits[1].Bit2;
OutputArray^.PDOs[24].6 := SignalArray.Segment3Color1Intensity.Bits[1].Bit3;

//Segment3 Animation Type
OutputArray^.PDOs[23].0 := SignalArray.Segment3AnimationType.Bits[1].Bit1;
OutputArray^.PDOs[23].1 := SignalArray.Segment3AnimationType.Bits[1].Bit2;
OutputArray^.PDOs[23].2 := SignalArray.Segment3AnimationType.Bits[1].Bit3;

//Segment 3 Speed
OutputArray^.PDOs[23].3 := SignalArray.Segment3Speed.Bits[1].Bit1;
OutputArray^.PDOs[23].4 := SignalArray.Segment3Speed.Bits[1].Bit2;

//Segment 3 Pulse Pattern
OutputArray^.PDOs[23].5 := SignalArray.Segment3PulsePattern.Bits[1].Bit1;
OutputArray^.PDOs[23].6 := SignalArray.Segment3PulsePattern.Bits[1].Bit2;

//Segment 3 Rotate
OutputArray^.PDOs[22].7 := SignalArray.Segment3RotationDir;

//Segment 3 Color 2
OutputArray^.PDOs[22].0 := SignalArray.Segment3Color2.Bits[1].Bit1;
OutputArray^.PDOs[22].1 := SignalArray.Segment3Color2.Bits[1].Bit2;
OutputArray^.PDOs[22].2 := SignalArray.Segment3Color2.Bits[1].Bit3;
OutputArray^.PDOs[22].3 := SignalArray.Segment3Color2.Bits[1].Bit4;

//Segment 3 Color 2 Intensity
OutputArray^.PDOs[22].4 := SignalArray.Segment3Color2Intensity.Bits[1].Bit1;
OutputArray^.PDOs[22].5 := SignalArray.Segment3Color2Intensity.Bits[1].Bit2;
OutputArray^.PDOs[22].6 := SignalArray.Segment3Color2Intensity.Bits[1].Bit3;
END_METHOD

END_FUNCTION_BLOCK

// ---- POUs/FBs/Devices/fb_Dev_StripLight_BannerWLS15Pro.TcPOU
(*
    fb_Dev_StripLight_BannerWLS15Pro
    ================================
    Drives a Banner WLS15 Pro RGB LED strip light (WLS15PXRGB<length>DSKQP)
    over IO-Link with the device in Run Mode -- Operating Mode Selection
    (index 0x40) = 1, which is how the light ships and how it is configured on
    this machine. Run Mode drives the WHOLE strip as one; use Segment Mode if
    independently addressable zones are ever needed.

    Run Mode carries one enumerated BYTE per parameter, so there is no
    sub-byte packing to do here -- unlike the TL50 Pro, whose fields are 1-4
    bits wide and share octets.

    The device's process data out is 32 bytes and Run Mode uses only the odd
    octets 13, 15, 17, 19, 21, 23, 25, 27, 29 and 31; the even octets are
    unused padding. A TwinCAT IO-Link port configured from the IODD publishes
    those ten as individually named port variables, so the PLC sees ten
    contiguous bytes and TwinCAT places them in the process image. That is why
    ST_Banner_WLS15PXRGB0220DSKQP_RunMode_Outputs is ten bytes and not
    thirty-two.

    Usage
    -----
        // IO.TcGVL -- link each member to the matching IO-Link port variable
        FIO2109_BannerLight AT %Q* : ST_Banner_WLS15PXRGB0220DSKQP_RunMode_Outputs;

        // Devices.TcGVL
        StripLight : fb_Dev_StripLight_BannerWLS15Pro(
                         cfgDeviceName     := 'Cell Strip Light',
                         cfgEnable         := TRUE,
                         cfgInitEventClass := TRUE);

        // MAIN -- steady green while running
        StripLight(refPDO       := ADR(IO.FIO2109_BannerLight),
                   inpAnimation := E_BannerWLS15Pro_Animation.eSteady,
                   inpColor1    := E_BannerWLS15Pro_Color.eGreen);

    The struct members are declared in the order TwinCAT lists the port
    variables, so they link straight down the list:
        Direction, Percent Width of Color 1, Scroll/Bounce Style,
        Color 2 Intensity, Color 2, Pulse Pattern, Speed,
        Color 1 Intensity, Color 1, Animation

    Reference: Banner "WLS15 Pro IO-Link Data Reference Guide", 219132 Rev. A,
    section 1.3.2 Run Mode.
*)
FUNCTION_BLOCK fb_Dev_StripLight_BannerWLS15Pro EXTENDS abs_fb_Device
VAR_INPUT
    // Process data out of the IO-Link port the light hangs off.
    refPDO                  : POINTER TO ST_Banner_WLS15PXRGB0220DSKQP_RunMode_Outputs;

    inpAnimation            : E_BannerWLS15Pro_Animation        := E_BannerWLS15Pro_Animation.eOff;
    inpColor1               : E_BannerWLS15Pro_Color            := E_BannerWLS15Pro_Color.eGreen;
    inpColor1Intensity      : E_BannerWLS15Pro_Intensity        := E_BannerWLS15Pro_Intensity.eHigh;
    inpColor2               : E_BannerWLS15Pro_Color            := E_BannerWLS15Pro_Color.eGreen;
    inpColor2Intensity      : E_BannerWLS15Pro_Intensity        := E_BannerWLS15Pro_Intensity.eHigh;
    inpSpeed                : E_BannerWLS15Pro_Speed            := E_BannerWLS15Pro_Speed.eMedium;
    // Only read by the flashing animations.
    inpPulsePattern         : E_BannerWLS15Pro_PulsePattern     := E_BannerWLS15Pro_PulsePattern.eNormal;
    // Only read by Scroll and Bounce.
    inpScrollBounceStyle    : E_BannerWLS15Pro_ScrollBounceStyle := E_BannerWLS15Pro_ScrollBounceStyle.eSolid;
    // Share of the strip lit with Color 1, in percent. The device accepts
    // 1..100 only, so this is clamped. Read by the Ends, Scroll and Bounce
    // animations; ignored by the rest.
    inpPercentWidthColor1   : BYTE                              := 50;
    inpDirection            : E_BannerWLS15Pro_Direction        := E_BannerWLS15Pro_Direction.eUp;
END_VAR

VAR_OUTPUT
    // FALSE means refPDO was never wired and nothing is reaching the light.
    stsLinked   : BOOL;
    // The value set last written, for readback and commissioning.
    stsShowing  : ST_Banner_WLS15PXRGB0220DSKQP_RunMode_Outputs;
END_VAR

VAR
    _out : ST_Banner_WLS15PXRGB0220DSKQP_RunMode_Outputs;
END_VAR

VAR CONSTANT
    cPERCENT_WIDTH_MIN : BYTE := 1;
    cPERCENT_WIDTH_MAX : BYTE := 100;
END_VAR

DeviceLogic();

// One enumerated byte per parameter -- the whole appearance is a value copy.
_out.Animnation             := TO_BYTE(inpAnimation);
_out.Color_1                := TO_BYTE(inpColor1);
_out.Color_1_Intensity      := TO_BYTE(inpColor1Intensity);
_out.Speed                  := TO_BYTE(inpSpeed);
_out.Pulse_Pattern          := TO_BYTE(inpPulsePattern);
_out.Color_2                := TO_BYTE(inpColor2);
_out.Color_2_Intensity      := TO_BYTE(inpColor2Intensity);
_out.Scroll_Bounce_Style    := TO_BYTE(inpScrollBounceStyle);
_out.Direction              := TO_BYTE(inpDirection);

// 0 and >100 are outside what the device accepts for the Color 1 width.
_out.Percent_Width_Of_Color_1 := LIMIT(cPERCENT_WIDTH_MIN, inpPercentWidthColor1, cPERCENT_WIDTH_MAX);

// A disabled or faulted light goes dark rather than holding its last pattern,
// so a stale display is never mistaken for a live one.
IF NOT _enabled OR stsFaulted THEN
    _out.Animnation := TO_BYTE(E_BannerWLS15Pro_Animation.eOff);
END_IF

stsLinked := (refPDO <> 0);

IF stsLinked THEN
    writeToPDO(inpValues := _out, inpTarget := refPDO);
END_IF

stsShowing := _out;

// Copies one Run Mode value set into the light's process data out.
METHOD PRIVATE writeToPDO : BOOL
VAR_INPUT
    inpValues : ST_Banner_WLS15PXRGB0220DSKQP_RunMode_Outputs;
    inpTarget : POINTER TO ST_Banner_WLS15PXRGB0220DSKQP_RunMode_Outputs;
END_VAR
// The octet numbers below are positions in the device's 32-byte Run Mode
// process image (219132 Rev. A, section 1.3.2). TwinCAT publishes each one as
// its own IO-Link port variable, so these members are linked one-to-one and
// the unused even octets never reach the PLC. Assigned member by member
// rather than as a whole-struct copy so a mis-ordered link is visible here.
inpTarget^.Direction                := inpValues.Direction;                 // octet 13
inpTarget^.Percent_Width_Of_Color_1 := inpValues.Percent_Width_Of_Color_1;  // octet 15
inpTarget^.Scroll_Bounce_Style      := inpValues.Scroll_Bounce_Style;       // octet 17
inpTarget^.Color_2_Intensity        := inpValues.Color_2_Intensity;         // octet 19
inpTarget^.Color_2                  := inpValues.Color_2;                   // octet 21
inpTarget^.Pulse_Pattern            := inpValues.Pulse_Pattern;             // octet 23
inpTarget^.Speed                    := inpValues.Speed;                     // octet 25
inpTarget^.Color_1_Intensity        := inpValues.Color_1_Intensity;         // octet 27
inpTarget^.Color_1                  := inpValues.Color_1;                   // octet 29
inpTarget^.Animnation               := inpValues.Animnation;                // octet 31

writeToPDO := TRUE;
END_METHOD

END_FUNCTION_BLOCK

// ---- POUs/FBs/Camming/fb_CamCoupler.TcPOU
// Reusable, machine-agnostic coupler: synchronizes ONE slave axis to a master axis via a verified
// NC cam table. Wraps MC_CamIn / MC_CamOut, gates engagement on the incoming
// 'verified' flag (from fb_CamTeach.stsVerified), coordinates the fb_Axis yield hook so the slave
// stops issuing its own motion while cammed, and decouples cleanly on fault/interlock loss.
//
// Standalone: does NOT extend abs_fb_Device. Its own error model (stsError/stsErrorText) is used
// instead of setFault, because a fault would gate the slave's MC_Power and break the coupling.
// Instantiate one per slave. The master is driven independently (elsewhere).
//
// NOTE ON INPUT NAMING: the design skeleton lists the couple/decouple triggers as VAR_INPUT
// 'cmdCouple'/'cmdDecouple'. Because this FB ALSO exposes public METHODS cmdCouple()/cmdDecouple()
// (both the input edges and the method calls start the sequences), the inputs are named inpCouple/
// inpDecouple to avoid an identifier collision - a method and a variable cannot share a name in
// TwinCAT. This matches the fb_Axis convention (inp* = wired inputs, cmd* = methods; cf. inpReset /
// cmdReset). Semantics are identical to the design skeleton. See report/deviations.
//
// THE TABLE: fb_CamTeach's download CREATES NC table 'tableId' (MC_CamTableSelect from the PLC
// points, periodicity fixed there) and verifies it; this coupler only engages that id with MC_CamIn.
// It does not select a table itself (an earlier MC_CamTableSelect here had no table data to give).
FUNCTION_BLOCK fb_CamCoupler
VAR_IN_OUT
    Master : AXIS_REF;                 // shared master (driven elsewhere)
    Slave  : AXIS_REF;                 // this slave
END_VAR

VAR_INPUT
    verified     : BOOL;               // from fb_CamTeach.stsVerified for this slave - REQUIRED to couple
    tableId      : UDINT;              // NC cam table id (same one fb_CamTeach downloaded); 0 = use cfgTableId
    periodic     : BOOL;               // informational (HMI echo): periodicity is set when fb_CamTeach creates the table
    masterOffset : LREAL;              // engage offsets to match current pose at master start
    slaveOffset  : LREAL;
    masterScale  : LREAL := 1.0;
    slaveScale   : LREAL := 1.0;
    interlockOK  : BOOL;               // machine/axis permissive
    slaveFB      : POINTER TO fb_Axis; // yield coordination (optional but recommended); 0 = no yield
    inpCouple    : BOOL;               // (design skeleton: cmdCouple) rising edge starts the couple sequence
    inpDecouple  : BOOL;               // (design skeleton: cmdDecouple) rising edge starts the decouple sequence
    inpReset     : BOOL;               // rising edge clears a latched error (back to E_CamCoupler_State.eIdle if safe)
END_VAR

VAR_OUTPUT
    stsCoupled   : BOOL;               // MC_CamIn.InSync
    stsBusy      : BOOL;               // a couple/decouple sequence is running
    stsState     : E_CamCoupler_State;
    stsError     : BOOL;               // latched coupler error (own model - not setFault)
    stsErrorText : STRING;
END_VAR

VAR
    // Public HMI interface - the struct an HMI (e.g. lhmi) binds
    HMI        : ST_CamCoupler_HMI_Interface;

    // MC camming / stop function blocks (Tc2_MC2 / Tc2_MC2_Camming)
    _camIn     : MC_CamIn;             // VERIFY against installed Tc2_MC2 / TF5050 version
    _camOut    : MC_CamOut;            // VERIFY against installed Tc2_MC2 / TF5050 version
    _mcHalt    : MC_Halt;              // stop the freed slave after CamOut
    _superImp  : MC_MoveSuperImposed;  // VERIFY against installed Tc2_MC2 / TF5050 version (live trim)

    _state : E_CamCoupler_State;       // working state (mirrored to stsState)

    // Command requests + input edge detectors
    _coupleReq    : BOOL;
    _decoupleReq  : BOOL;
    _resetReq     : BOOL;
    _trigCouple   : R_TRIG;
    _trigDecouple : R_TRIG;
    _trigReset    : R_TRIG;

    // Sequence control flags
    _engaged       : BOOL;             // in one of the engaged states (yielding..coupled)
    _beginDecouple : BOOL;             // request to start the decouple path this scan
    _faultDecouple : BOOL;             // TRUE = the active decouple was fault-triggered (end in E_CamCoupler_State.eError)
    _slaveReady    : BOOL;             // slave powered/operational (best-effort via AXIS_REF + slaveFB)
    _camInExec     : BOOL;             // MC_CamIn.Execute driver (TRUE from eCoupling through eCoupled)
    _camInRetrig   : INT;              // 0=idle, 1=drop Execute one scan, 2=re-execute (live offset trim)
    _haltExec      : BOOL;             // MC_Halt.Execute driver (post-CamOut stop)

    // Superimposed correction (live trim)
    _superImpReq   : BOOL;             // one-shot start request
    _superImpExec  : BOOL;             // MC_MoveSuperImposed.Execute driver
    _superImpDist  : LREAL;
    _superImpVelo  : LREAL;
    _superImpAccel : LREAL := 100.0;   // [slave unit/s2] accel/decel for the corrective move

    // Effective engage parameters (resolved from inputs/cfg at couple; latched so live trim persists)
    _tableId      : UDINT;
    _periodic     : BOOL;
    _masterOffset : LREAL;
    _slaveOffset  : LREAL;
    _masterScale  : LREAL := 1.0;
    _slaveScale   : LREAL := 1.0;

    // Commissioning defaults (FB_Init / cfg* properties)
    _cfgTableId   : UDINT;
    _cfgPeriodic  : BOOL;

    // Stop dynamics for the post-CamOut halt
    _haltDecel    : LREAL := 100.0;    // [slave unit/s2]

    _hmiCfgLoaded : BOOL;              // HMI.Config seeded from defaults once
END_VAR

// ── 1. Refresh AXIS_REF status snapshots ─────────────────────────────────────
// Decode NcToPlc into Master/Slave .Status before anything reads .Status this scan. fb_Axis refreshes
// the same shared refs each scan; a second ReadStatus() here is harmless and keeps this FB self-contained.
Master.ReadStatus();
Slave.ReadStatus();

// Slave "enabled / operational" check. Best-effort via the shared AXIS_REF, refined by the slave's
// fb_Axis power state when the pointer is wired. (Pointer deref guarded - IEC OR/AND do not short-circuit.)
_slaveReady := (NOT Slave.Status.Disabled) AND (NOT Slave.Status.ErrorStop) AND (NOT Slave.Status.Error);
IF slaveFB <> 0 THEN
    _slaveReady := _slaveReady AND slaveFB^.stsEnabled;
END_IF

// ── 2. Command inputs: rising edges + self-clearing HMI one-shots ─────────────
// Both the wired input edges and the public methods funnel into the same request flags.
_trigCouple(CLK := inpCouple);
IF _trigCouple.Q THEN cmdCouple(); END_IF
_trigDecouple(CLK := inpDecouple);
IF _trigDecouple.Q THEN cmdDecouple(); END_IF
_trigReset(CLK := inpReset);
IF _trigReset.Q THEN cmdReset(); END_IF

IF HMI.Commands.ocmdCouple THEN
    HMI.Commands.ocmdCouple := FALSE;
    cmdCouple();
END_IF
IF HMI.Commands.ocmdDecouple THEN
    HMI.Commands.ocmdDecouple := FALSE;
    cmdDecouple();
END_IF
IF HMI.Commands.ocmdReset THEN
    HMI.Commands.ocmdReset := FALSE;
    cmdReset();
END_IF
IF HMI.Commands.ocmdSetMasterOffset THEN
    HMI.Commands.ocmdSetMasterOffset := FALSE;
    cmdSetMasterOffset(HMI.Commands.ocmdMasterOffset);
END_IF
IF HMI.Commands.ocmdSetSlaveOffset THEN
    HMI.Commands.ocmdSetSlaveOffset := FALSE;
    cmdSetSlaveOffset(HMI.Commands.ocmdSlaveOffset);
END_IF
IF HMI.Commands.ocmdSuperImpose THEN
    HMI.Commands.ocmdSuperImpose := FALSE;
    cmdSuperImpose(HMI.Commands.ocmdSuperImposeDist, HMI.Commands.ocmdSuperImposeVelo);
END_IF

// ── 3. Reset ─────────────────────────────────────────────────────────────────
// Honored only from a resting state - a reset must never tear down an active coupling.
IF _resetReq THEN
    _resetReq := FALSE;
    IF _state = E_CamCoupler_State.eError OR _state = E_CamCoupler_State.eIdle THEN
        stsError       := FALSE;
        stsErrorText   := '';
        _faultDecouple := FALSE;
        _state         := E_CamCoupler_State.eIdle;
    END_IF
END_IF

// ── 4. Safety & decouple triggers ────────────────────────────────────────────
// Evaluated BEFORE the state machine so a loss condition begins the decouple the same scan it appears.
_engaged := (_state = eYielding) OR (_state = eSelecting) OR (_state = eCoupling) OR (_state = eCoupled);
_beginDecouple := FALSE;

// Operator-requested decouple (only meaningful while engaged).
IF _decoupleReq THEN
    _decoupleReq := FALSE;
    IF _engaged THEN
        _faultDecouple := FALSE;
        _beginDecouple := TRUE;
    END_IF
END_IF

// Fault / interlock loss / verified drop while engaged -> forced decouple + latched error.
// No auto re-couple: a deliberate cmdCouple (after a reset) is required to re-engage.
// MC_CamIn is hard-gated on verified below, so a dropped 'verified' both aborts and prevents re-engage.
IF _engaged AND NOT stsError THEN
    IF NOT interlockOK THEN
        raiseError('Interlock lost while coupled');
        _faultDecouple := TRUE;
        _beginDecouple := TRUE;
    ELSIF Slave.Status.Error THEN
        raiseError(CONCAT('Slave axis error: ', UDINT_TO_STRING(Slave.NcToPlc.ErrorCode)));
        _faultDecouple := TRUE;
        _beginDecouple := TRUE;
    ELSIF NOT verified THEN
        raiseError('Verified dropped while coupled');
        _faultDecouple := TRUE;
        _beginDecouple := TRUE;
    END_IF
END_IF

IF _beginDecouple THEN
    _camInExec := FALSE;
    IF _camIn.InSync OR (_state = eCoupled) OR (_state = eCoupling) THEN
        _state := eDecoupling;         // disengage the cam first (CamOut)
    ELSE
        _haltExec := TRUE;
        _state    := eStopping;        // not cammed yet - just stop the slave & release the yield
    END_IF
END_IF

// ── 5. Couple / decouple state machine ───────────────────────────────────────
CASE _state OF

    E_CamCoupler_State.eIdle:
        _camInExec := FALSE;
        _haltExec  := FALSE;
        IF _coupleReq THEN
            _coupleReq := FALSE;
            // Preconditions (design: verified, slave enabled, interlockOK, not already coupled).
            IF NOT verified THEN
                raiseError('Cannot couple: table not verified');
                _state := E_CamCoupler_State.eError;
            ELSIF NOT interlockOK THEN
                raiseError('Cannot couple: interlock not OK');
                _state := E_CamCoupler_State.eError;
            ELSIF _camIn.InSync THEN
                raiseError('Cannot couple: already coupled');
                _state := E_CamCoupler_State.eError;
            ELSIF NOT _slaveReady THEN
                raiseError('Cannot couple: slave not enabled');
                _state := E_CamCoupler_State.eError;
            ELSE
                // Resolve effective table id / periodicity (live input overrides the commissioning
                // default; periodic input is authoritative - the machine layer supplies it per slave).
                IF tableId <> 0 THEN _tableId := tableId; ELSE _tableId := _cfgTableId; END_IF
                _periodic := periodic;
                // Yield: fb_Axis runs an interruptible halt, then suppresses all its own motion.
                IF slaveFB <> 0 THEN
                    slaveFB^.cmdSetExternalControl(TRUE);
                END_IF
                _state := eYielding;
            END_IF
        END_IF

    eYielding:
        // Wait for the slave to reach standstill (the fb_Axis entry cmdHalt completes) before engaging,
        // so the halt and the coupling never overlap (design coupler note). The table already exists
        // (fb_CamTeach created + verified it), so engage straight away.
        IF Slave.Status.Standstill THEN
            // Latch engage parameters from the inputs at engage time (so later live trim persists).
            _masterOffset := masterOffset;
            _slaveOffset  := slaveOffset;
            IF masterScale <> 0.0 THEN _masterScale := masterScale; ELSE _masterScale := 1.0; END_IF
            IF slaveScale  <> 0.0 THEN _slaveScale  := slaveScale;  ELSE _slaveScale  := 1.0; END_IF
            _camInExec := TRUE;        // begin engaging
            _state     := eCoupling;
        END_IF

    eCoupling:
        // MC_CamIn driven Execute:=_camInExec (section 7). Engage complete when InSync.
        IF _camIn.InSync THEN
            _state := eCoupled;
        ELSIF _camIn.Error THEN
            raiseError(CONCAT('CamIn error: ', UDINT_TO_STRING(_camIn.ErrorID)));
            _camInExec     := FALSE;
            _faultDecouple := TRUE;
            _state         := eDecoupling;   // CamOut to be safe, then stop -> E_CamCoupler_State.eError
        ELSIF _camIn.CommandAborted THEN
            raiseError('CamIn aborted');
            _camInExec     := FALSE;
            _faultDecouple := TRUE;
            _state         := eDecoupling;
        END_IF

    eCoupled:
        // Steady state - coupling held. Live trim (offset re-issue / superimpose) runs in sections 7 & 10.
        // External loss conditions are handled in section 4; an NC-level CamIn error is caught here.
        IF _camIn.Error THEN
            raiseError(CONCAT('CamIn error: ', UDINT_TO_STRING(_camIn.ErrorID)));
            _camInExec     := FALSE;
            _faultDecouple := TRUE;
            _state         := eDecoupling;
        END_IF

    eDecoupling:
        // MC_CamOut driven Execute:=TRUE by state gate (section 8).
        IF _camOut.Done THEN
            _haltExec := TRUE;         // slave keeps its last velocity after CamOut -> halt it
            _state    := eStopping;
        ELSIF _camOut.Error THEN
            raiseError(CONCAT('CamOut error: ', UDINT_TO_STRING(_camOut.ErrorID)));
            _faultDecouple := TRUE;
            _haltExec      := TRUE;    // still try to bring the slave to rest & release the yield
            _state         := eStopping;
        END_IF

    eStopping:
        // MC_Halt driven Execute:=_haltExec (section 9). Done when at rest.
        IF _mcHalt.Done OR Slave.Status.Standstill THEN
            _haltExec := FALSE;
            // Release the yield: fb_Axis resumes control and stays at rest until a new explicit command.
            IF slaveFB <> 0 THEN
                slaveFB^.cmdSetExternalControl(FALSE);
            END_IF
            IF _faultDecouple THEN
                _faultDecouple := FALSE;
                _state         := E_CamCoupler_State.eError;   // stsError already latched by raiseError
            ELSE
                _state := E_CamCoupler_State.eIdle;
            END_IF
        END_IF

    E_CamCoupler_State.eError:
        // Latched fault - wait for cmdReset/inpReset. No motion commanded here.
        _camInExec := FALSE;
        _haltExec  := FALSE;

END_CASE

// ── 6. (no table select - fb_CamTeach created the table; see the header) ─────

// ── 7. MC_CamIn (engage - RampIn, offset/scaling) ────────────────────────────
// Live offset trim re-issues MC_CamIn: drop Execute for one scan, then re-execute with the new offsets.
IF _camInRetrig = 1 THEN
    _camInExec   := FALSE;
    _camInRetrig := 2;
ELSIF _camInRetrig = 2 THEN
    _camInExec   := TRUE;
    _camInRetrig := 0;
END_IF
// HARD gate on 'verified': never engage an unverified table (design principle 2).
// VERIFY against installed Tc2_MC2 / TF5050 version: StartMode enum name/values (RampIn variant),
// CamTableID type (MC_CAM_ID) and source, and MasterOffset/SlaveOffset/MasterScaling/SlaveScaling
// semantics + which StartMode supports live offset re-issue.
_camIn(
    Master        := Master,
    Slave         := Slave,
    Execute       := _camInExec AND verified,
    MasterOffset  := _masterOffset,
    SlaveOffset   := _slaveOffset,
    MasterScaling := _masterScale,
    SlaveScaling  := _slaveScale,
    StartMode     := MC_STARTMODE_ABSOLUTE,    // absolute: cam CS congruent with axis CS (no RampIn member in this TF5050)
    CamTableID    := _tableId                   // the table fb_CamTeach created and verified
);

// ── 8. MC_CamOut (disengage) ─────────────────────────────────────────────────
// VERIFY against installed Tc2_MC2 / TF5050 version: block signature (Slave-only in/out).
_camOut(
    Slave   := Slave,
    Execute := (_state = eDecoupling)
);

// ── 9. MC_Halt (kill the retained slave velocity after CamOut) ───────────────
_mcHalt(
    Axis         := Slave,
    Execute      := _haltExec,
    Deceleration := _haltDecel,
    Jerk         := 0.0
);
IF _mcHalt.Done THEN
    _haltExec := FALSE;
END_IF

// ── 10. MC_MoveSuperImposed (live corrective move on top of the cam) ──────────
// Kept engaged: a bounded correction superimposed on the running cam (no decouple).
IF _superImpReq THEN
    _superImpReq  := FALSE;
    _superImpExec := TRUE;
END_IF
// VERIFY against installed Tc2_MC2 / TF5050 version: block signature and VelocityDiff semantics
// (superimposed on a synchronized/cammed axis).
_superImp(
    Axis         := Slave,
    Execute      := _superImpExec,
    Distance     := _superImpDist,
    VelocityDiff := _superImpVelo,
    Acceleration := _superImpAccel,
    Deceleration := _superImpAccel,
    Jerk         := 0.0
);
IF _superImp.Done OR _superImp.CommandAborted OR _superImp.Error THEN
    _superImpExec := FALSE;
END_IF

// ── 11. Outputs ──────────────────────────────────────────────────────────────
stsState   := _state;
stsCoupled := _camIn.InSync;
stsBusy    := (_state = eYielding) OR (_state = eSelecting) OR (_state = eCoupling)
              OR (_state = eDecoupling) OR (_state = eStopping);

// ── 12. HMI status update ────────────────────────────────────────────────────
// Seed the commissioning mirror once from the configured defaults.
IF NOT _hmiCfgLoaded THEN
    HMI.Config.tableId      := _cfgTableId;
    HMI.Config.periodic     := _cfgPeriodic;
    HMI.Config.masterOffset := _masterOffset;
    HMI.Config.slaveOffset  := _slaveOffset;
    HMI.Config.masterScale  := _masterScale;
    HMI.Config.slaveScale   := _slaveScale;
    _hmiCfgLoaded := TRUE;
END_IF
HMI.Status.stsState        := _state;
HMI.Status.stsCoupled      := stsCoupled;
HMI.Status.stsBusy         := stsBusy;
HMI.Status.stsError        := stsError;
HMI.Status.stsErrorText    := stsErrorText;
HMI.Status.stsVerified     := verified;
HMI.Status.stsTableId      := _tableId;
HMI.Status.stsMasterOffset := _masterOffset;
HMI.Status.stsSlaveOffset  := _slaveOffset;
HMI.Status.stsMasterScale  := _masterScale;
HMI.Status.stsSlaveScale   := _slaveScale;
HMI.Status.stsPeriodic     := _periodic;

// Request an engage of this slave onto the master via the verified cam table.
// Multi-scan sequence: yield -> select -> cam-in. Accepted only from E_CamCoupler_State.eIdle; rejected QUIETLY while
// busy/engaged/errored (no fault - a fault would gate the slave MC_Power and break any coupling).
// Reachable both from this method and the rising edge of inpCouple.
METHOD PUBLIC cmdCouple : BOOL
IF _state <> E_CamCoupler_State.eIdle THEN
    cmdCouple := FALSE;
    RETURN;
END_IF

_coupleReq := TRUE;
cmdCouple  := TRUE;
END_METHOD

// Request a controlled decouple: CamOut -> MC_Halt (kill retained velocity) -> release the yield.
// Ignored QUIETLY if not engaged. Reachable both from this method and the rising edge of inpDecouple.
METHOD PUBLIC cmdDecouple : BOOL
_decoupleReq := TRUE;
cmdDecouple  := TRUE;
END_METHOD

// Clear a latched coupler error and return to E_CamCoupler_State.eIdle. Honored only from E_CamCoupler_State.eError/E_CamCoupler_State.eIdle so it can never
// tear down an active coupling. Reachable from this method, ocmdReset, and the rising edge of inpReset.
METHOD PUBLIC cmdReset : BOOL
_resetReq := TRUE;
cmdReset  := TRUE;
END_METHOD

// Live master-offset trim (no decouple): re-issue MC_CamIn with the new master offset while the
// coupling stays engaged. Accepted only while fully coupled; rejected QUIETLY otherwise.
METHOD PUBLIC cmdSetMasterOffset : BOOL
VAR_INPUT
    offset : LREAL;   // [master unit] new cam master offset
END_VAR
IF _state <> eCoupled THEN
    cmdSetMasterOffset := FALSE;
    RETURN;
END_IF

_masterOffset      := offset;
_camInRetrig       := 1;   // one clear scan, then MC_CamIn re-executes with the new offset
cmdSetMasterOffset := TRUE;
END_METHOD

// Live slave-offset trim (no decouple): re-issue MC_CamIn with the new slave offset while the
// coupling stays engaged. Accepted only while fully coupled; rejected QUIETLY otherwise.
METHOD PUBLIC cmdSetSlaveOffset : BOOL
VAR_INPUT
    offset : LREAL;   // [slave unit] new cam slave offset
END_VAR
IF _state <> eCoupled THEN
    cmdSetSlaveOffset := FALSE;
    RETURN;
END_IF

_slaveOffset      := offset;
_camInRetrig      := 1;   // one clear scan, then MC_CamIn re-executes with the new offset
cmdSetSlaveOffset := TRUE;
END_METHOD

// Bounded corrective move superimposed on top of the running cam via MC_MoveSuperImposed (no decouple).
// Accepted only while fully coupled and no correction is already active; rejected QUIETLY otherwise.
METHOD PUBLIC cmdSuperImpose : BOOL
VAR_INPUT
    distance : LREAL;   // [slave unit] corrective distance added on top of the cam
    velocity : LREAL;   // [slave unit/s] additional velocity for the correction
END_VAR
IF _state <> eCoupled THEN
    cmdSuperImpose := FALSE;
    RETURN;
END_IF

IF _superImpExec THEN
    // one correction at a time
    cmdSuperImpose := FALSE;
    RETURN;
END_IF

_superImpDist  := distance;
_superImpVelo  := velocity;
_superImpReq   := TRUE;    // rising-edge Execute in section 10 next scan
cmdSuperImpose := TRUE;
END_METHOD

// Latch the FB's own error. This FB does NOT extend abs_fb_Device and deliberately does NOT call
// setFault: a fault would gate the slave MC_Power and drop the coupling. Preserves the first cause
// if several conditions trip in the same scan.
METHOD PRIVATE raiseError : BOOL
VAR_INPUT
    text : STRING;
END_VAR
IF NOT stsError THEN
    stsError     := TRUE;
    stsErrorText := text;
END_IF
raiseError := TRUE;
END_METHOD

// Return the full HMI interface struct (the one an HMI binds).
METHOD PUBLIC getHMIdata : ST_CamCoupler_HMI_Interface
getHMIdata := HMI;
END_METHOD

METHOD FB_Init : BOOL
VAR_INPUT
    bInitRetains : BOOL;
    bInCopyCode  : BOOL;
    cfgTableId   : UDINT;   // commissioning default NC cam table id
    cfgPeriodic  : BOOL;    // commissioning default periodicity
END_VAR
THIS^._cfgTableId  := cfgTableId;
THIS^._cfgPeriodic := cfgPeriodic;
// Seed the effective values so status/HMI reflect the defaults before the first couple.
THIS^._tableId  := cfgTableId;
THIS^._periodic := cfgPeriodic;
END_METHOD

// Commissioning default NC cam table id, used when the tableId VAR_INPUT is left 0.
PROPERTY PUBLIC cfgTableId : UDINT
GET
cfgTableId := _cfgTableId;
END_GET
SET
_cfgTableId := cfgTableId;
END_SET
END_PROPERTY

// Commissioning default periodicity. The periodic VAR_INPUT is authoritative at couple time; this
// seeds the power-on default for setups that drive the coupler without wiring that input.
PROPERTY PUBLIC cfgPeriodic : BOOL
GET
cfgPeriodic := _cfgPeriodic;
END_GET
SET
_cfgPeriodic := cfgPeriodic;
END_SET
END_PROPERTY

END_FUNCTION_BLOCK

// ---- POUs/FBs/fb_Axis.TcPOU
// Single-axis wrapper. Extends abs_fb_Device for fault/interlock/event infrastructure.
// Axis-level interlocks are set externally via cmdSetInterlock (inherited).
// Move-level interlocks live in each move's ST_Interlock field; a parallel array of
// fb_Interlock instances (one per slot) evaluates them every scan.
FUNCTION_BLOCK fb_Axis EXTENDS abs_fb_Device
VAR_INPUT
    // Inherited from abs_fb_Device:
    //   inpAuto            : BOOL  -- machine in automatic mode
    //   inpReset           : BOOL  -- machine-level reset (resets axis)
    //   inpInterlockBypass : BOOL  -- bypass axis-level interlock
    //   faultMonitor       : POINTER TO fb_FaultMonitor
    inpSTO  : BOOL;     // Safe Torque Off feedback - TRUE = STO not active (normal), FALSE = STO active
                        // Safety program provides ~350ms between STP drop and STO activation.
                        // Falling edge immediately triggers MC_Stop for graceful decel in that window.
    // Global velocity override (machine-wide). Wire from a machine-level source (e.g. a shared
    // GVL) so one control can drive many axes. When inpGlobalOverrideEnable is TRUE the effective
    // velocity override is inpGlobalOverride [%]; otherwise the axis-local override set from the
    // HMI. Reported via stsVelocityOverride (effective value) + stsGlobalOverrideActive.
    inpGlobalOverrideEnable : BOOL;   // TRUE = follow the global override; FALSE = use local
    inpGlobalOverride       : INT;    // [%] global velocity override, clamped 0..100 (0 = axis held)

    // Physical teach-pendant jog (hardware-wired, level-triggered like the HMI jog). Same safety
    // gating and arbitration as HMI jog, but driven by MC_MoveVelocity (section 12b), NOT _mcJog:
    // MC_Jog takes its speed once, at the jog's start, so a stick pushed further or B pressed
    // mid-jog did nothing - and the start fired as the stick crossed the activation threshold, so
    // every jog latched whatever deflection that instant had. Never two motion sources at once. The pendant OWNS the jog while it is selected (inpPendantMode) or its dead-man is
    // held (inpPendantEnable): the HMI jog, torque-jog and go-to are locked out, so the two can't
    // command opposite directions. Motion still needs the dead-man. Manual mode only, same as HMI
    // jog. Reported via HMI.Status.stsJogSource / stsPendantMode / stsPendantDeadman.
    inpPendantMode     : BOOL;    // pendant selected - locks out HMI jog even before the dead-man is held
    inpPendantEnable   : BOOL;    // dead-man / enable - must be held for pendant jog (and to take ownership)
    inpPendantJogPos   : BOOL;    // jog forward  (level: held = jog)
    inpPendantJogNeg   : BOOL;    // jog backward (level: held = jog)
    inpPendantJogVelo  : LREAL;   // [unit/s]  pendant jog velocity     (<= 0 = use configured jog velocity)
    inpPendantJogAccel : LREAL;   // [unit/s²] pendant jog acceleration (<= 0 = use configured jog accel)
    inpPendantJogFraction : LREAL; // 0..1 of the pendant base speed (inpPendantJogVelo if > 0, else the
                                   // configured jog speed) AFTER the NC-max clamp, so full deflection is
                                   // exactly the axis's top jog speed. <= 0 = not used (base speed as-is).
                                   // Follows live: stick / speed-modifier changes apply mid-jog.
END_VAR

VAR_IN_OUT
    Axis  : AXIS_REF;
END_VAR

VAR_OUTPUT
    stsEnabled    : BOOL;   // drive powered (MC_Power.Status)
    stsMoving     : BOOL;   // axis in motion
    stsStandstill : BOOL;   // powered and at rest
    stsInTarget   : BOOL;   // within position target window
    stsMoveDone   : BOOL;   // last position/velocity move reached setpoint
    stsCurrentMove: INT;    // index of current/last executed move (0 = none)
    // Live process values, also exposed as direct outputs (not just via HMI.Status) so the
    // calling program can wire them to charts / data logging / other logic. Sourced from Axis.NcToPlc.
    stsActualPosition : LREAL;   // [unit]   actual position (Axis.NcToPlc.ActPos)
    stsActualVelocity : LREAL;   // [unit/s] actual velocity (Axis.NcToPlc.ActVelo)
    stsActualTorque   : LREAL;   // [% or Nm] actual torque (Axis.NcToPlc.ActTorque)
    stsNcMaxVelocity  : LREAL;   // [unit/s] the NC axis's maximum velocity (MC_ReadParameterSet; 0 until read)
    // Setpoints (paired with the actuals above). Position/velocity come from the NC
    // setpoint generator (Axis.NcToPlc.Set*). There is NO NC torque setpoint — torque is
    // commanded straight to the drive — so stsSetTorque is the torque this FB is commanding
    // (active move's torque, torque-jog value, or 0).
    stsSetPosition    : LREAL;   // [unit]   commanded position (Axis.NcToPlc.SetPos)
    stsSetVelocity    : LREAL;   // [unit/s] commanded velocity (Axis.NcToPlc.SetVelo)
    stsSetTorque      : LREAL;   // [% or Nm] commanded torque (FB-tracked; no NC setpoint exists)
END_VAR

VAR
    // Public HMI interface - the struct an HMI (e.g. lhmi) binds
    HMI             : ST_Axis_HMI_Interface;

    // Per-move interlock FBs (parallel to moves array; cannot embed FB in struct)
    _moveInterlocks : ARRAY[1..20] OF fb_Interlock;

    // MC Function Blocks
    _mcPower        : MC_Power;
    _mcReset        : MC_Reset;
    _mcStop         : MC_Stop;
    _mcHalt         : MC_Halt;
    _mcMoveAbs      : MC_MoveAbsolute;
    _mcMoveRel      : MC_MoveRelative;
    _mcMoveVel      : MC_MoveVelocity;
    _mcMoveMod      : MC_MoveModulo;     // eModulo: absolute target WITHIN one modulo period, forced direction
    _mcReadParams   : MC_ReadParameterSet;  // the NC axis parameter set: fVeloMaximum clamps jog speeds (section 12)
    _mcTorque       : MC_TorqueControl;     // Tc2_MC2 torque mode with continuous setpoint updates
    _mcTorqueJog    : MC_TorqueControl;     // dedicated instance for interactive torque-jog (dead-man)
    _mcJog          : MC_Jog;           // HMI jog only (the pendant uses _mcPendantVel / _mcPendantHalt)
    _mcPendantVel   : MC_MoveVelocity;  // pendant jog: re-triggered when the speed changes (section 12b)
    _mcPendantHalt  : MC_Halt;          // pendant jog release: ramp to standstill at the jog accel
    _mcHome         : MC_Home;          // MC_Direct: sets position only (does NOT set calibrated flag)
    _mcForceCal     : MC_Home;          // MC_ForceCalibration: sets the calibrated/Homed flag without moving
    _mcOverride     : MC_SetOverride;
    _mcJogGoto      : MC_MoveAbsolute;   // position jog ("go to position") - dedicated instance, section 12c
    _mcRestorePos   : MC_SetPosition;    // retained home: re-applies the stored offset after an NC restart (10b)
    _mcRestoreCal   : MC_Home;           // retained home: MC_ForceCalibration after the restore (10b)

    // Internal state
    _isEnabled          : BOOL;
    _externalControl    : BOOL;
    _currentMoveIndex   : INT;
    _activeMoveMode     : E_Axis_Mode;
    _moveExecState      : INT;          // 0=idle, 1=abort-scan, 2=executing
    _startMoveReq       : BOOL;
    _pendingIndex       : INT;
    _pendingMode        : E_Axis_Mode;

    _stopCmd            : BOOL;         // MC_Stop active - locked until cmdReset
    _haltCmd            : BOOL;         // MC_Halt active - auto-clears on done
    _resetCmd           : BOOL;
    _homeCmd            : BOOL;
    _homeStep           : INT;          // 0=idle, 1=MC_Direct (set pos), 2=MC_ForceCalibration (set Homed)
    _homePosition       : LREAL;

    // --- Home diagnostics: MC_Direct/MC_ForceCalibration finish in ~1 scan (no motion),
    //     so Done/Busy/Active pulses are invisible online. These LATCH so you can eyeball
    //     what happened after a home. All reset at the start of each cmdHome. ---
    _dbgHomeMaxStep     : INT;          // highest _homeStep reached (want 2)
    _dbgHomeDirectDone  : BOOL;         // MC_Direct (step 1) reported Done
    _dbgHomeCalDone     : BOOL;         // MC_ForceCalibration (step 2) reported Done
    _dbgHomeCalError    : BOOL;         // MC_ForceCalibration reported Error
    _dbgHomeCalErrID    : UDINT;        // ...its ErrorID

    _jogPositive        : BOOL;
    _jogNegative        : BOOL;
    _jogVelocity        : LREAL := 10.0;
    _jogAccel           : LREAL := 100.0;
    _jogSource          : E_Axis_JogSource;    // which input owns the jog this scan (HMI vs pendant)
    _jogVeloEff         : LREAL := 10.0;        // effective jog velocity fed to _mcJog (pendant speed when it owns; else _jogVelocity)
    _jogAccelEff        : LREAL := 100.0;       // effective jog accel    fed to _mcJog
    _ncMaxVelocity      : LREAL;                // [unit/s] NC max velocity (0 = not read yet -> no clamp)
    _axisParams         : ST_AxisParameterSet;  // MC_ReadParameterSet target
    _readParamsExec     : BOOL;
    _readParamsRetry    : TON;                  // (re)try the read every 2 s until it succeeds
    _lastMcErrorId      : UDINT;                // last motion-block error (jog/move/home) - published as stsErrorID
    _jogErrorEdge       : R_TRIG;               // MC_Jog.Error rising edge -> fault (was silent)
    // Pendant jog (section 12b)
    _pjGate             : BOOL;                 // the jog safety gate (same terms as MC_Jog's JogForward/Backwards)
    _pjDir              : INT;                  // this scan: 1 forward, -1 backward, 0 none
    _pjDirPrev          : INT;
    _pjVelExec          : BOOL;                 // _mcPendantVel.Execute
    _pjVeloSent         : LREAL;                // [unit/s] speed latched into the running MC_MoveVelocity
    _pjRetrig           : TON;                  // min time between speed re-triggers
    _pjMoving           : BOOL;                 // a pendant velocity command was issued and has not been halted yet
    _pjErrorEdge        : R_TRIG;
    // Position jog ("go to position"): discrete absolute move, jog subvariant (see section 12c).
    _jogGotoTarget      : LREAL;            // [unit] operator-entered absolute target (angle or mm)
    _jogGotoBusy        : BOOL;             // go-to move in progress - mutually exclusive with jog / moves / home
    _jogTorqueLimit     : LREAL;            // [Nm or %] global overtorque trip for position jog (0 = no limit).
                                            //   Exceed → locked MC_Stop + fault 'Overtorque limit: jog'.
                                            //   Applies to position jog only; torque-jog is bounded by _torqueJogMaxLimit.

    // Torque jog (dead-man interactive torque). Held → command the entered torque; released
    // → command 0 (ramps down) and disengage once actual torque ~0 (stays enabled, no MC_Stop).
    _torqueJogActive    : BOOL;             // button held this scan (gated) → apply torque
    _torqueJogEngaged   : BOOL;             // block active: held, or ramping back to 0 after release
    _torqueJogValue     : LREAL;            // clamped live torque setpoint [% rated]
    _torqueJogRamp      : LREAL := 500.0;   // [% rated/s] ramp for torque changes / release
    _torqueJogMaxLimit  : LREAL := 100.0;   // [% rated] absolute clamp on the entered torque
    _tjMaxVelInit       : BOOL;             // FALSE until the retained _tjMaxVel is echoed to the HMI once (re-armed each restart)

    _velocityOverride   : LREAL := 100.0;   // [%] 0-100 (axis-local, set from HMI)
    _accelOverride      : LREAL := 100.0;   // [%] 0-100
    _activeVelocityOverride : LREAL := 100.0;   // [%] effective override actually applied (global if enabled, else local)
    _stopDecel          : LREAL := 1000.0;  // [unit/s²] decel for MC_Stop
    _haltDecel          : LREAL := 100.0;   // [unit/s²] decel for MC_Halt

    // [% rated] |ActTorque| below this = torque released → torque-jog disengages
    // (see section 12b). Also the "torque is back to ~0" threshold after a released dead-man.
    _stopTorqueThreshold : LREAL := 1.0;

    _axisType           : E_Axis_UnitType := E_Axis_UnitType.eLinear;  // HMI: linear vs rotary
    _unit               : STRING := 'mm';   // HMI position unit label (velocity = unit + '/s')
    // TRUE = the NC axis is configured as modulo. NC config carries no runtime "modulo on/off"
    // flag in the cyclic image, so it's declared here (like _axisType/_unit). Drives which
    // position the HMI shows: modulo (Axis.NcToPlc.ModuloActPos, wrapped into one period) vs the
    // accumulated Axis.NcToPlc.ActPos. Orthogonal to _axisType — a rotary axis need not be modulo.
    _isModulo           : BOOL;

    _selectedMove       : INT;          // HMI move staged for confirmation
    _confirmPending     : BOOL;
    _hmiMoveConfigLoaded: BOOL;
    _moveConfigApplyError: BOOL;
    _moveConfigErrorText : STRING;

    _stoFallingEdge     : F_TRIG;       // detects STO drop for graceful stop initiation

    _i                  : INT;          // loop index
    _moveConfigValid    : BOOL;

    // Retained operator settings / home (see VAR PERSISTENT, sections 1b and 10b)
    _settingsInit       : BOOL;         // FALSE until the retained settings are applied + echoed to the HMI (once per start)
    _lastHmiJogVelocity : LREAL;        // HMI field last scan - an operator edit is a CHANGE of the field
    _lastHmiJogAccel    : LREAL;
    _retainHome         : BOOL := TRUE; // see cfgRetainHome
    _homeActAtStart     : LREAL;        // [unit] ActPos captured when a teach starts
    _ncOffsetApplied    : LREAL;        // [unit] offset the RUNNING NC currently applies to the raw encoder position
    _homeRestoreChecked : BOOL;         // the once-per-start retained-home check has run
    _homeRestoreDelay   : TON;          // axis IO must be valid this long before the check runs
    _homeRestoreStep    : INT;          // 0=idle, 1=MC_SetPosition, 2=MC_ForceCalibration
    _homeRestoreTarget  : LREAL;        // [unit] raw position + retained offset
END_VAR

VAR PERSISTENT
    // FB-owned live move table. HMI.Config.moves is an edit buffer; accepted
    // edits are copied here and retained with the fb_Axis instance.
    moves : ARRAY[1..20] OF ST_Axis_MoveDefinition;
    // Torque-jog overspeed trip [unit/s], 0 = off. Retained across restart; edited live
    // from HMI.Commands.ocmdTorqueJogMaxVel (see the torque-jog section, ~12b).
    _tjMaxVel : LREAL;
    // Operator jog / override settings. 0 = never set by an operator → the FB_Init/cfg default
    // stands. Applied over the defaults once per start (section 1b), so they survive a restart.
    _savedJogVelocity      : LREAL;     // [unit/s]
    _savedJogAccel         : LREAL;     // [unit/s²]
    _savedVelocityOverride : LREAL;     // [%] 0 < x <= 100
    // Taught home, kept until the next teach (section 10b): taught position = raw encoder
    // position + _homeOffset. Needs an absolute encoder.
    _homeTaught    : BOOL;
    _homeOffset    : LREAL;             // [unit]
    _homeTaughtPos : LREAL;             // [unit] the position that was taught (HMI display)
END_VAR

// ── 1. Base device logic ─────────────────────────────────────────────────────
// Processes axis-level interlock, raises/clears fault events, updates HMIbasedevice.
// Also calls cmdReset() if inpReset is TRUE (machine reset resets axis).
DeviceLogic();

// Refresh the decoded AXIS_REF.Status snapshot from the cyclic NcToPlc data BEFORE
// anything reads Axis.Status.* this scan. Without this, Status fields (notably
// .Homed/calibrated) can lag the real NC state even though the NC faceplate shows
// it correctly — Status is only guaranteed current right after ReadStatus().
Axis.ReadStatus();

// ── 1b. Retained operator settings ────────────────────────────────────────────
// FB_Init re-seeds jog velocity/accel from the instance declaration on every cold start, and
// HMI.Commands is plain VAR, so without this an activation reset the operator's values. Once per
// start, lay the retained values (VAR PERSISTENT) over the defaults and echo them to the HMI
// fields so the HMI shows them instead of re-sending its power-up zeros. Edits are retained as
// they are entered (section 3).
IF NOT _settingsInit THEN
    IF _savedJogVelocity > 0.0 THEN
        _jogVelocity := _savedJogVelocity;
    END_IF
    IF _savedJogAccel > 0.0 THEN
        _jogAccel := _savedJogAccel;
    END_IF
    IF _savedVelocityOverride > 0.0 AND _savedVelocityOverride <= 100.0 THEN
        _velocityOverride := _savedVelocityOverride;
    END_IF
    IF _homeTaught THEN
        _homePosition           := _homeTaughtPos;
        HMI.Config.homePosition := _homeTaughtPos;
    END_IF
    HMI.Commands.ocmdJogVelocity      := _jogVelocity;
    HMI.Commands.ocmdJogAcceleration  := _jogAccel;
    HMI.Commands.ocmdVelocityOverride := _velocityOverride;
    _lastHmiJogVelocity := _jogVelocity;
    _lastHmiJogAccel    := _jogAccel;
    _settingsInit := TRUE;
END_IF

// ── 2. Evaluate all move interlocks each scan ─────────────────────────────────
FOR _i := 1 TO 20 DO
    _moveInterlocks[_i].name := CONCAT(moves[_i].moveName, '_ILK');
    _moveInterlocks[_i](inpConfig := moves[_i].interlock);
END_FOR

IF NOT _hmiMoveConfigLoaded THEN
    FOR _i := 1 TO 20 DO
        HMI.Config.moves[_i] := moves[_i];
    END_FOR
    _hmiMoveConfigLoaded := TRUE;
END_IF

// ── 3. HMI commands ───────────────────────────────────────────────────────────
// Reset is accepted in both auto and manual.
IF HMI.Commands.ocmdReset THEN
    HMI.Commands.ocmdReset := FALSE;
    cmdReset();
END_IF

IF NOT _inAuto THEN

    IF HMI.Commands.ocmdEnable THEN
        HMI.Commands.ocmdEnable := FALSE;
        cmdEnable();
    END_IF

    IF HMI.Commands.ocmdDisable THEN
        HMI.Commands.ocmdDisable := FALSE;
        cmdDisable();
    END_IF

    IF HMI.Commands.ocmdStop THEN
        HMI.Commands.ocmdStop := FALSE;
        cmdStop();
    END_IF

    IF HMI.Commands.ocmdHome THEN
        HMI.Commands.ocmdHome := FALSE;
        cmdHome(HMI.Config.homePosition);
    END_IF

    // Position jog ("go to position"): run a discrete absolute move to the entered target.
    // Locked out (quietly) while the teach pendant owns the jog, like the HMI jog buttons.
    IF HMI.Commands.ocmdJogGoto THEN
        HMI.Commands.ocmdJogGoto := FALSE;
        IF NOT inpPendantMode AND NOT inpPendantEnable THEN
            cmdJogGoto(HMI.Commands.ocmdJogGotoPos);
        END_IF
    END_IF

    // Move selection: two-step - select then confirm
    IF HMI.Commands.ocmdSelectMove >= 1 AND HMI.Commands.ocmdSelectMove <= 20 THEN
        _selectedMove   := HMI.Commands.ocmdSelectMove;
        _confirmPending := TRUE;
        HMI.Commands.ocmdSelectMove := 0;
    END_IF

    IF HMI.Commands.ocmdCancelSelect THEN
        HMI.Commands.ocmdCancelSelect := FALSE;
        _selectedMove   := 0;
        _confirmPending := FALSE;
    END_IF

    IF HMI.Commands.ocmdReloadMoveConfig THEN
        HMI.Commands.ocmdReloadMoveConfig := FALSE;
        FOR _i := 1 TO 20 DO
            HMI.Config.moves[_i] := moves[_i];
        END_FOR
        _moveConfigApplyError := FALSE;
        _moveConfigErrorText  := '';
    END_IF

    IF HMI.Commands.ocmdApplyMoveConfig THEN
        HMI.Commands.ocmdApplyMoveConfig := FALSE;

        IF _moveExecState <> 0 OR Axis.Status.DiscreteMotion OR Axis.Status.ContinuousMotion OR Axis.Status.Stopping THEN
            _moveConfigApplyError := TRUE;
            _moveConfigErrorText  := 'Cannot apply move config while axis is active';
        ELSE
            _moveConfigValid := TRUE;
            _moveConfigErrorText := '';

            FOR _i := 1 TO 20 DO
                IF HMI.Config.moves[_i].velocity < 0.0 THEN
                    _moveConfigValid := FALSE;
                    _moveConfigErrorText := CONCAT('Move velocity < 0 at index ', INT_TO_STRING(_i));
                ELSIF HMI.Config.moves[_i].acceleration < 0.0 THEN
                    _moveConfigValid := FALSE;
                    _moveConfigErrorText := CONCAT('Move acceleration < 0 at index ', INT_TO_STRING(_i));
                ELSIF HMI.Config.moves[_i].deceleration < 0.0 THEN
                    _moveConfigValid := FALSE;
                    _moveConfigErrorText := CONCAT('Move deceleration < 0 at index ', INT_TO_STRING(_i));
                ELSIF HMI.Config.moves[_i].jerk < 0.0 THEN
                    _moveConfigValid := FALSE;
                    _moveConfigErrorText := CONCAT('Move jerk < 0 at index ', INT_TO_STRING(_i));
                ELSIF HMI.Config.moves[_i].torqueRamp < 0.0 THEN
                    _moveConfigValid := FALSE;
                    _moveConfigErrorText := CONCAT('Move torque ramp < 0 at index ', INT_TO_STRING(_i));
                ELSIF HMI.Config.moves[_i].cfgTorqueLimit < 0.0 THEN
                    _moveConfigValid := FALSE;
                    _moveConfigErrorText := CONCAT('Move torque limit < 0 at index ', INT_TO_STRING(_i));
                END_IF
            END_FOR

            IF _moveConfigValid THEN
                FOR _i := 1 TO 20 DO
                    moves[_i] := HMI.Config.moves[_i];
                END_FOR
                _selectedMove := 0;
                _confirmPending := FALSE;
                _moveConfigApplyError := FALSE;
                _moveConfigErrorText  := '';
            ELSE
                _moveConfigApplyError := TRUE;
            END_IF
        END_IF
    END_IF

    // Always self-clear ocmdRunMove when seen — otherwise a Run pressed with nothing staged
    // (or after reset/disable cleared _confirmPending) latches TRUE and auto-fires the NEXT
    // Select. Only actually start a move when one is staged.
    IF HMI.Commands.ocmdRunMove THEN
        HMI.Commands.ocmdRunMove := FALSE;
        IF _confirmPending THEN
            _confirmPending := FALSE;
            cmdStart(_selectedMove);
        END_IF
    END_IF

    // Jog arbitration: physical teach pendant vs HMI. Level-triggered - hold to jog. Both feed the
    // ONE _mcJog (section 12); they are never two motion sources. The pendant OWNS the jog from the
    // moment it is selected (inpPendantMode) or its dead-man is held (inpPendantEnable): the HMI jog
    // buttons are ignored, so the two can't fight over direction. Pendant motion still needs the
    // dead-man. Within a source, forward AND backward together is contradictory -> no request (no
    // motion). Blocked while homing / mid-move / torque-jogging.
    IF _externalControl OR _jogGotoBusy THEN
        // Yielded to a coordinator (e.g. fb_CamCoupler) or a go-to move is running - no speed jog.
        _jogSource   := E_Axis_JogSource.eNone;
        _jogPositive := FALSE;
        _jogNegative := FALSE;
    ELSIF inpPendantMode OR inpPendantEnable THEN
        _jogSource   := E_Axis_JogSource.ePendant;
        _jogPositive := inpPendantEnable AND inpPendantJogPos AND NOT inpPendantJogNeg AND NOT _homeCmd AND (_moveExecState = 0);
        _jogNegative := inpPendantEnable AND inpPendantJogNeg AND NOT inpPendantJogPos AND NOT _homeCmd AND (_moveExecState = 0);
    ELSIF HMI.Commands.ocmdJogPositive AND NOT HMI.Commands.ocmdJogNegative AND NOT HMI.Commands.ocmdTorqueJog AND NOT _homeCmd AND (_moveExecState = 0) THEN
        _jogSource   := E_Axis_JogSource.eHMI;
        _jogVelocity := SEL(HMI.Commands.ocmdJogVelocity     > 0.0, _jogVelocity, HMI.Commands.ocmdJogVelocity);
        _jogAccel    := SEL(HMI.Commands.ocmdJogAcceleration > 0.0, _jogAccel,    HMI.Commands.ocmdJogAcceleration);
        _jogPositive := TRUE;
        _jogNegative := FALSE;
    ELSIF HMI.Commands.ocmdJogNegative AND NOT HMI.Commands.ocmdJogPositive AND NOT HMI.Commands.ocmdTorqueJog AND NOT _homeCmd AND (_moveExecState = 0) THEN
        _jogSource   := E_Axis_JogSource.eHMI;
        _jogVelocity := SEL(HMI.Commands.ocmdJogVelocity     > 0.0, _jogVelocity, HMI.Commands.ocmdJogVelocity);
        _jogAccel    := SEL(HMI.Commands.ocmdJogAcceleration > 0.0, _jogAccel,    HMI.Commands.ocmdJogAcceleration);
        _jogNegative := TRUE;
        _jogPositive := FALSE;
    ELSE
        _jogSource   := E_Axis_JogSource.eNone;
        _jogPositive := FALSE;
        _jogNegative := FALSE;
    END_IF

    // Torque jog: dead-man. Held = command the entered torque; gated the same as jog
    // (no home, no running move, no position jog, not while the pendant owns the jog).
    // Release/engage + ramp handled in section 12b.
    _torqueJogActive := HMI.Commands.ocmdTorqueJog
        AND NOT _externalControl AND NOT _jogGotoBusy
        AND NOT _jogPositive AND NOT _jogNegative
        AND NOT inpPendantMode AND NOT inpPendantEnable
        AND NOT _homeCmd AND (_moveExecState = 0);
    IF _torqueJogActive THEN
        _torqueJogValue := LIMIT(-_torqueJogMaxLimit, HMI.Commands.ocmdTorqueJogValue, _torqueJogMaxLimit);
    END_IF

    // Operator settings take effect - and are retained (section 1b) - as soon as they are entered,
    // not only on the next HMI jog press, so an edit survives a restart even if it was never used.
    // Jog velocity/accel are adopted on an HMI EDIT (field changed since last scan), so a value set
    // from PLC code (cfgJog* property, cmdJog* argument) is not reverted by a stale HMI field.
    IF HMI.Commands.ocmdJogVelocity > 0.0 AND HMI.Commands.ocmdJogVelocity <> _lastHmiJogVelocity THEN
        _jogVelocity      := HMI.Commands.ocmdJogVelocity;
        _savedJogVelocity := _jogVelocity;
    END_IF
    _lastHmiJogVelocity := HMI.Commands.ocmdJogVelocity;
    IF HMI.Commands.ocmdJogAcceleration > 0.0 AND HMI.Commands.ocmdJogAcceleration <> _lastHmiJogAccel THEN
        _jogAccel      := HMI.Commands.ocmdJogAcceleration;
        _savedJogAccel := _jogAccel;
    END_IF
    _lastHmiJogAccel := HMI.Commands.ocmdJogAcceleration;
    IF HMI.Commands.ocmdVelocityOverride > 0.0 AND HMI.Commands.ocmdVelocityOverride <= 100.0 THEN
        _velocityOverride      := HMI.Commands.ocmdVelocityOverride;
        _savedVelocityOverride := _velocityOverride;
    END_IF

ELSE
    // AUTO: no operator jogging. The jog arbitration above runs only in manual, so a jog or
    // torque-jog button held across the manual -> auto switch would otherwise stay latched and
    // keep the axis jogging (or applying torque) in Auto. Drop any jog an OPERATOR source owns;
    // a jog started by PLC code through cmdJogPositive/cmdJogNegative has _jogSource = eNone and
    // is left alone. Torque jog is operator-only, so it always stops (section 12b ramps it to 0).
    IF _jogSource <> E_Axis_JogSource.eNone THEN
        _jogSource   := E_Axis_JogSource.eNone;
        _jogPositive := FALSE;
        _jogNegative := FALSE;
    END_IF
    _torqueJogActive := FALSE;
END_IF

// ── 4. STO handling ──────────────────────────────────────────────────────────
// STO active (inpSTO FALSE) is treated as a SOFT operational inhibit, not a fault:
// MC_Power.Enable is gated by inpSTO at the level (section 6) so the drive can't be
// powered while STO is active, and stsSafetyInhibited annunciates it. A semi-auto
// sequence can open the guard, do a manual step, close it, and resume WITHOUT a reset.
//
// A fault is raised ONLY when STO drops while the axis was actually moving/commanded —
// an uncommanded stop mid-motion must be acknowledged. In that case fire MC_Stop for a
// graceful decel within the ~350ms window before hardware cuts torque, and latch a fault
// (cleared by a deliberate cmdReset). No automatic restart: pending moves are always
// dropped here, so motion never resumes on its own — a new cmdStart is required either way.
_stoFallingEdge(CLK := inpSTO);
IF _stoFallingEdge.Q THEN
    // Cancel any pending / held motion commands regardless of case.
    _haltCmd       := FALSE;
    _jogPositive   := FALSE;
    _jogNegative   := FALSE;
    _homeCmd       := FALSE;
    _startMoveReq  := FALSE;
    _jogGotoBusy   := FALSE;
    // Abnormal only: was moving / mid-move / applying torque → graceful stop + latched fault.
    // (Jog and position moves show up as NC Discrete/ContinuousMotion; torque paths via
    // _moveExecState / _torqueJogEngaged.) Evaluate BEFORE zeroing _moveExecState below.
    IF    Axis.Status.DiscreteMotion OR Axis.Status.ContinuousMotion OR Axis.Status.Stopping
       OR (_moveExecState <> 0) OR _torqueJogEngaged THEN
        _stopCmd := TRUE;
        setFault(TRUE, 'STO during motion');
    END_IF
    _moveExecState := 0;
END_IF

// ── 5. Axis interlock loss during motion → forced stop ────────────────────────
// Safety event: use MC_Stop (locked standstill, not interruptible).
IF _mcPower.Status AND NOT Interlock.outInterlockOK THEN
    IF Axis.Status.DiscreteMotion OR Axis.Status.ContinuousMotion OR Axis.Status.Stopping THEN
        _stopCmd       := TRUE;
        _haltCmd       := FALSE;
        _jogPositive   := FALSE;
        _jogNegative   := FALSE;
        _homeCmd       := FALSE;
        _startMoveReq  := FALSE;
        _jogGotoBusy   := FALSE;
        _moveExecState := 0;
        IF NOT stsFaulted THEN
            setFault(TRUE, CONCAT('I_NOK during motion: ', Interlock.stsFirstOut));
        END_IF
    END_IF
END_IF

// ── 6. MC_Power ───────────────────────────────────────────────────────────────
// inpSTO gates Enable at the level: drive cannot be powered while STO is active,
// regardless of software enable state or fault clear.
_mcPower(
    Axis            := Axis,
    Enable          := _isEnabled AND NOT stsFaulted AND inpSTO,
    Enable_Positive := TRUE,
    Enable_Negative := TRUE,
    Override        := 1.0,
    BufferMode      := 0
);

// ── 7. MC_Reset ───────────────────────────────────────────────────────────────
_mcReset(Axis := Axis, Execute := _resetCmd);
IF _mcReset.Done OR _mcReset.Error THEN
    _resetCmd := FALSE;
END_IF

// ── 8. MC_Stop (forced standstill) ───────────────────────────────────────────
// _stopCmd remains TRUE until cmdReset clears it.
_mcStop(
    Axis         := Axis,
    Execute      := _stopCmd,
    Deceleration := _stopDecel,
    Jerk         := 0.0
);

// ── 9. MC_Halt (interruptible stop) ──────────────────────────────────────────
// Auto-clears when standstill reached; new cmdStart can resume. Also clears when the halt is
// superseded (CommandAborted) or refused (Error): _haltCmd used to stay TRUE then, so the NEXT
// cmdHalt found Execute already high, produced no rising edge and halted NOTHING - an axis handed
// back from external control kept running at its last commanded speed.
_mcHalt(
    Axis         := Axis,
    Execute      := _haltCmd,
    Deceleration := _haltDecel,
    Jerk         := 0.0
);
IF _mcHalt.Done OR _mcHalt.CommandAborted OR _mcHalt.Error THEN
    _haltCmd := FALSE;
END_IF

